       "DB_Bad_Konfig".Bad_Konfig[1].IO_Ein.WT_Einsetzen[1] := "FB_KP8_DB_1".KP8.Taste[6];
       "DB_Bad_Konfig".Bad_Konfig[1].IO_Ein.WT_Einsetzen[2] := "FB_KP8_DB_1".KP8.Taste[5];
       "DB_Bad_Konfig".Bad_Konfig[1].IO_Ein.WT_Einsetzen[3] := "FB_KP8_DB_1".KP8.Taste[4];
       "DB_Bad_Konfig".Bad_Konfig[1].IO_Ein.WT_Entnehmen[1] := "FB_KP8_DB_1".KP8.Taste[2];
       "DB_Bad_Konfig".Bad_Konfig[1].IO_Ein.WT_Entnehmen[2] := "FB_KP8_DB_1".KP8.Taste[1];
       "DB_Bad_Konfig".Bad_Konfig[1].IO_Ein.WT_Entnehmen[3] := "FB_KP8_DB_1".KP8.Taste[0];
       "DB_Bad_Konfig".Bad_Konfig[3].IO_Ein.WT_Einsetzen[1] := "FB_KP8_DB_2".KP8.Taste[6];
       "DB_Bad_Konfig".Bad_Konfig[3].IO_Ein.WT_Einsetzen[2] := "FB_KP8_DB_2".KP8.Taste[5];
       "DB_Bad_Konfig".Bad_Konfig[3].IO_Ein.WT_Einsetzen[3] := "FB_KP8_DB_2".KP8.Taste[4];
       "DB_Bad_Konfig".Bad_Konfig[3].IO_Ein.WT_Entnehmen[1] := "FB_KP8_DB_2".KP8.Taste[2];
       "DB_Bad_Konfig".Bad_Konfig[3].IO_Ein.WT_Entnehmen[2] := "FB_KP8_DB_2".KP8.Taste[1];
       "DB_Bad_Konfig".Bad_Konfig[3].IO_Ein.WT_Entnehmen[3] := "FB_KP8_DB_2".KP8.Taste[0];
       "DB_Bad_Konfig".Bad_Konfig[7].IO_Ein.WT_Einsetzen[1] := "FB_KP8_DB_4".KP8.Taste[6];
       "DB_Bad_Konfig".Bad_Konfig[7].IO_Ein.WT_Einsetzen[2] := "FB_KP8_DB_4".KP8.Taste[5];
       "DB_Bad_Konfig".Bad_Konfig[7].IO_Ein.WT_Einsetzen[3] := "FB_KP8_DB_4".KP8.Taste[4];
       "DB_Bad_Konfig".Bad_Konfig[7].IO_Ein.WT_Entnehmen[1] := "FB_KP8_DB_4".KP8.Taste[2];
       "DB_Bad_Konfig".Bad_Konfig[7].IO_Ein.WT_Entnehmen[2] := "FB_KP8_DB_4".KP8.Taste[1];
       "DB_Bad_Konfig".Bad_Konfig[7].IO_Ein.WT_Entnehmen[3] := "FB_KP8_DB_4".KP8.Taste[0];
       "DB_Bad_Konfig".Bad_Konfig[8].IO_Ein.WT_Einsetzen[1] := "FB_KP8_DB_5".KP8.Taste[6];
       "DB_Bad_Konfig".Bad_Konfig[8].IO_Ein.WT_Einsetzen[2] := "FB_KP8_DB_5".KP8.Taste[5];
       "DB_Bad_Konfig".Bad_Konfig[8].IO_Ein.WT_Einsetzen[3] := "FB_KP8_DB_5".KP8.Taste[4];
       "DB_Bad_Konfig".Bad_Konfig[8].IO_Ein.WT_Entnehmen[1] := "FB_KP8_DB_5".KP8.Taste[2];
       "DB_Bad_Konfig".Bad_Konfig[8].IO_Ein.WT_Entnehmen[2] := "FB_KP8_DB_5".KP8.Taste[1];
       "DB_Bad_Konfig".Bad_Konfig[8].IO_Ein.WT_Entnehmen[3] := "FB_KP8_DB_5".KP8.Taste[0];
       "DB_Bad_Konfig".Bad_Konfig[12].IO_Ein.WT_Einsetzen[1] := "FB_KP8_DB_7".KP8.Taste[6];
       "DB_Bad_Konfig".Bad_Konfig[12].IO_Ein.WT_Einsetzen[2] := "FB_KP8_DB_7".KP8.Taste[5];
       "DB_Bad_Konfig".Bad_Konfig[12].IO_Ein.WT_Einsetzen[3] := "FB_KP8_DB_7".KP8.Taste[4];
       "DB_Bad_Konfig".Bad_Konfig[12].IO_Ein.WT_Entnehmen[1] := "FB_KP8_DB_7".KP8.Taste[2];
       "DB_Bad_Konfig".Bad_Konfig[12].IO_Ein.WT_Entnehmen[2] := "FB_KP8_DB_7".KP8.Taste[1];
       "DB_Bad_Konfig".Bad_Konfig[12].IO_Ein.WT_Entnehmen[3] := "FB_KP8_DB_7".KP8.Taste[0];
       "DB_Bad_Konfig".Bad_Konfig[13].IO_Ein.WT_Einsetzen[1] := "FB_KP8_DB_8".KP8.Taste[6];
       "DB_Bad_Konfig".Bad_Konfig[13].IO_Ein.WT_Einsetzen[2] := "FB_KP8_DB_8".KP8.Taste[5];
       "DB_Bad_Konfig".Bad_Konfig[13].IO_Ein.WT_Einsetzen[3] := "FB_KP8_DB_8".KP8.Taste[4];
       "DB_Bad_Konfig".Bad_Konfig[13].IO_Ein.WT_Entnehmen[1] := "FB_KP8_DB_8".KP8.Taste[2];
       "DB_Bad_Konfig".Bad_Konfig[13].IO_Ein.WT_Entnehmen[2] := "FB_KP8_DB_8".KP8.Taste[1];
       "DB_Bad_Konfig".Bad_Konfig[13].IO_Ein.WT_Entnehmen[3] := "FB_KP8_DB_8".KP8.Taste[0];
       "DB_Bad_Konfig".Bad_Konfig[14].IO_Ein.WT_Einsetzen[1] := "FB_KP8_DB_9".KP8.Taste[6];
       "DB_Bad_Konfig".Bad_Konfig[14].IO_Ein.WT_Einsetzen[2] := "FB_KP8_DB_9".KP8.Taste[5];
       "DB_Bad_Konfig".Bad_Konfig[14].IO_Ein.WT_Einsetzen[3] := "FB_KP8_DB_9".KP8.Taste[4];
       "DB_Bad_Konfig".Bad_Konfig[14].IO_Ein.WT_Entnehmen[1] := "FB_KP8_DB_9".KP8.Taste[2];
       "DB_Bad_Konfig".Bad_Konfig[14].IO_Ein.WT_Entnehmen[2] := "FB_KP8_DB_9".KP8.Taste[1];
       "DB_Bad_Konfig".Bad_Konfig[14].IO_Ein.WT_Entnehmen[3] := "FB_KP8_DB_9".KP8.Taste[0];
       "DB_Bad_Konfig".Bad_Konfig[18].IO_Ein.WT_Einsetzen[1] := "FB_KP8_DB_11".KP8.Taste[6];
       "DB_Bad_Konfig".Bad_Konfig[18].IO_Ein.WT_Einsetzen[2] := "FB_KP8_DB_11".KP8.Taste[5];
       "DB_Bad_Konfig".Bad_Konfig[18].IO_Ein.WT_Einsetzen[3] := "FB_KP8_DB_11".KP8.Taste[4];
       "DB_Bad_Konfig".Bad_Konfig[18].IO_Ein.WT_Entnehmen[1] := "FB_KP8_DB_11".KP8.Taste[2];
       "DB_Bad_Konfig".Bad_Konfig[18].IO_Ein.WT_Entnehmen[2] := "FB_KP8_DB_11".KP8.Taste[1];
       "DB_Bad_Konfig".Bad_Konfig[18].IO_Ein.WT_Entnehmen[3] := "FB_KP8_DB_11".KP8.Taste[0];
       "DB_Bad_Konfig".Bad_Konfig[19].IO_Ein.WT_Einsetzen[1] := "FB_KP8_DB_12".KP8.Taste[6];
       "DB_Bad_Konfig".Bad_Konfig[19].IO_Ein.WT_Einsetzen[2] := "FB_KP8_DB_12".KP8.Taste[5];
       "DB_Bad_Konfig".Bad_Konfig[19].IO_Ein.WT_Einsetzen[3] := "FB_KP8_DB_12".KP8.Taste[4];
       "DB_Bad_Konfig".Bad_Konfig[19].IO_Ein.WT_Entnehmen[1] := "FB_KP8_DB_12".KP8.Taste[2];
       "DB_Bad_Konfig".Bad_Konfig[19].IO_Ein.WT_Entnehmen[2] := "FB_KP8_DB_12".KP8.Taste[1];
       "DB_Bad_Konfig".Bad_Konfig[19].IO_Ein.WT_Entnehmen[3] := "FB_KP8_DB_12".KP8.Taste[0];
       "DB_Bad_Konfig".Bad_Konfig[21].IO_Ein.WT_Einsetzen[1] := "FB_KP8_DB_13".KP8.Taste[6];
       "DB_Bad_Konfig".Bad_Konfig[21].IO_Ein.WT_Einsetzen[2] := "FB_KP8_DB_13".KP8.Taste[5];
       "DB_Bad_Konfig".Bad_Konfig[21].IO_Ein.WT_Einsetzen[3] := "FB_KP8_DB_13".KP8.Taste[4];
       "DB_Bad_Konfig".Bad_Konfig[21].IO_Ein.WT_Entnehmen[1] := "FB_KP8_DB_13".KP8.Taste[2];
       "DB_Bad_Konfig".Bad_Konfig[21].IO_Ein.WT_Entnehmen[2] := "FB_KP8_DB_13".KP8.Taste[1];
       "DB_Bad_Konfig".Bad_Konfig[21].IO_Ein.WT_Entnehmen[3] := "FB_KP8_DB_13".KP8.Taste[0];
       "DB_Bad_Konfig".Bad_Konfig[26].IO_Ein.WT_Einsetzen[1] := "FB_KP8_DB_15".KP8.Taste[6];
       "DB_Bad_Konfig".Bad_Konfig[26].IO_Ein.WT_Einsetzen[2] := "FB_KP8_DB_15".KP8.Taste[5];
       "DB_Bad_Konfig".Bad_Konfig[26].IO_Ein.WT_Einsetzen[3] := "FB_KP8_DB_15".KP8.Taste[4];
       "DB_Bad_Konfig".Bad_Konfig[26].IO_Ein.WT_Entnehmen[1] := "FB_KP8_DB_15".KP8.Taste[2];
       "DB_Bad_Konfig".Bad_Konfig[26].IO_Ein.WT_Entnehmen[2] := "FB_KP8_DB_15".KP8.Taste[1];
       "DB_Bad_Konfig".Bad_Konfig[26].IO_Ein.WT_Entnehmen[3] := "FB_KP8_DB_15".KP8.Taste[0];
       "DB_Bad_Konfig".Bad_Konfig[30].IO_Ein.WT_Einsetzen[1] := "FB_KP8_DB_17".KP8.Taste[6];
       "DB_Bad_Konfig".Bad_Konfig[30].IO_Ein.WT_Einsetzen[2] := "FB_KP8_DB_17".KP8.Taste[5];
       "DB_Bad_Konfig".Bad_Konfig[30].IO_Ein.WT_Einsetzen[3] := "FB_KP8_DB_17".KP8.Taste[4];
       "DB_Bad_Konfig".Bad_Konfig[30].IO_Ein.WT_Entnehmen[1] := "FB_KP8_DB_17".KP8.Taste[2];
       "DB_Bad_Konfig".Bad_Konfig[30].IO_Ein.WT_Entnehmen[2] := "FB_KP8_DB_17".KP8.Taste[1];
       "DB_Bad_Konfig".Bad_Konfig[30].IO_Ein.WT_Entnehmen[3] := "FB_KP8_DB_17".KP8.Taste[0];
       "DB_Bad_Konfig".Bad_Konfig[31].IO_Ein.WT_Einsetzen[1] := "FB_KP8_DB_18".KP8.Taste[6];
       "DB_Bad_Konfig".Bad_Konfig[31].IO_Ein.WT_Einsetzen[2] := "FB_KP8_DB_18".KP8.Taste[5];
       "DB_Bad_Konfig".Bad_Konfig[31].IO_Ein.WT_Einsetzen[3] := "FB_KP8_DB_18".KP8.Taste[4];
       "DB_Bad_Konfig".Bad_Konfig[31].IO_Ein.WT_Entnehmen[1] := "FB_KP8_DB_18".KP8.Taste[2];
       "DB_Bad_Konfig".Bad_Konfig[31].IO_Ein.WT_Entnehmen[2] := "FB_KP8_DB_18".KP8.Taste[1];
       "DB_Bad_Konfig".Bad_Konfig[31].IO_Ein.WT_Entnehmen[3] := "FB_KP8_DB_18".KP8.Taste[0];
       "DB_Bad_Konfig".Bad_Konfig[35].IO_Ein.WT_Einsetzen[1] := "FB_KP8_DB_20".KP8.Taste[6];
       "DB_Bad_Konfig".Bad_Konfig[35].IO_Ein.WT_Einsetzen[2] := "FB_KP8_DB_20".KP8.Taste[5];
       "DB_Bad_Konfig".Bad_Konfig[35].IO_Ein.WT_Einsetzen[3] := "FB_KP8_DB_20".KP8.Taste[4];
       "DB_Bad_Konfig".Bad_Konfig[35].IO_Ein.WT_Entnehmen[1] := "FB_KP8_DB_20".KP8.Taste[2];
       "DB_Bad_Konfig".Bad_Konfig[35].IO_Ein.WT_Entnehmen[2] := "FB_KP8_DB_20".KP8.Taste[1];
       "DB_Bad_Konfig".Bad_Konfig[35].IO_Ein.WT_Entnehmen[3] := "FB_KP8_DB_20".KP8.Taste[0];
       "DB_Bad_Konfig".Bad_Konfig[36].IO_Ein.WT_Einsetzen[1] := "FB_KP8_DB_21".KP8.Taste[6];
       "DB_Bad_Konfig".Bad_Konfig[36].IO_Ein.WT_Einsetzen[2] := "FB_KP8_DB_21".KP8.Taste[5];
       "DB_Bad_Konfig".Bad_Konfig[36].IO_Ein.WT_Einsetzen[3] := "FB_KP8_DB_21".KP8.Taste[4];
       "DB_Bad_Konfig".Bad_Konfig[36].IO_Ein.WT_Entnehmen[1] := "FB_KP8_DB_21".KP8.Taste[2];
       "DB_Bad_Konfig".Bad_Konfig[36].IO_Ein.WT_Entnehmen[2] := "FB_KP8_DB_21".KP8.Taste[1];
       "DB_Bad_Konfig".Bad_Konfig[36].IO_Ein.WT_Entnehmen[3] := "FB_KP8_DB_21".KP8.Taste[0];
       "DB_Bad_Konfig".Bad_Konfig[40].IO_Ein.WT_Einsetzen[1] := "FB_KP8_DB_23".KP8.Taste[6];
       "DB_Bad_Konfig".Bad_Konfig[40].IO_Ein.WT_Einsetzen[2] := "FB_KP8_DB_23".KP8.Taste[5];
       "DB_Bad_Konfig".Bad_Konfig[40].IO_Ein.WT_Einsetzen[3] := "FB_KP8_DB_23".KP8.Taste[4];
       "DB_Bad_Konfig".Bad_Konfig[40].IO_Ein.WT_Entnehmen[1] := "FB_KP8_DB_23".KP8.Taste[2];
       "DB_Bad_Konfig".Bad_Konfig[40].IO_Ein.WT_Entnehmen[2] := "FB_KP8_DB_23".KP8.Taste[1];
       "DB_Bad_Konfig".Bad_Konfig[40].IO_Ein.WT_Entnehmen[3] := "FB_KP8_DB_23".KP8.Taste[0];
       "DB_Bad_Konfig".Bad_Konfig[41].IO_Ein.WT_Einsetzen[1] := "FB_KP8_DB_24".KP8.Taste[6];
       "DB_Bad_Konfig".Bad_Konfig[41].IO_Ein.WT_Einsetzen[2] := "FB_KP8_DB_24".KP8.Taste[5];
       "DB_Bad_Konfig".Bad_Konfig[41].IO_Ein.WT_Einsetzen[3] := "FB_KP8_DB_24".KP8.Taste[4];
       "DB_Bad_Konfig".Bad_Konfig[41].IO_Ein.WT_Entnehmen[1] := "FB_KP8_DB_24".KP8.Taste[2];
       "DB_Bad_Konfig".Bad_Konfig[41].IO_Ein.WT_Entnehmen[2] := "FB_KP8_DB_24".KP8.Taste[1];
       "DB_Bad_Konfig".Bad_Konfig[41].IO_Ein.WT_Entnehmen[3] := "FB_KP8_DB_24".KP8.Taste[0];
       "DB_Bad_Konfig".Bad_Konfig[45].IO_Ein.WT_Einsetzen[1] := "FB_KP8_DB_26".KP8.Taste[6];
       "DB_Bad_Konfig".Bad_Konfig[45].IO_Ein.WT_Einsetzen[2] := "FB_KP8_DB_26".KP8.Taste[5];
       "DB_Bad_Konfig".Bad_Konfig[45].IO_Ein.WT_Einsetzen[3] := "FB_KP8_DB_26".KP8.Taste[4];
       "DB_Bad_Konfig".Bad_Konfig[45].IO_Ein.WT_Entnehmen[1] := "FB_KP8_DB_26".KP8.Taste[2];
       "DB_Bad_Konfig".Bad_Konfig[45].IO_Ein.WT_Entnehmen[2] := "FB_KP8_DB_26".KP8.Taste[1];
       "DB_Bad_Konfig".Bad_Konfig[45].IO_Ein.WT_Entnehmen[3] := "FB_KP8_DB_26".KP8.Taste[0];
       "DB_Bad_Konfig".Bad_Konfig[46].IO_Ein.WT_Einsetzen[1] := "FB_KP8_DB_27".KP8.Taste[6];
       "DB_Bad_Konfig".Bad_Konfig[46].IO_Ein.WT_Einsetzen[2] := "FB_KP8_DB_27".KP8.Taste[5];
       "DB_Bad_Konfig".Bad_Konfig[46].IO_Ein.WT_Einsetzen[3] := "FB_KP8_DB_27".KP8.Taste[4];
       "DB_Bad_Konfig".Bad_Konfig[46].IO_Ein.WT_Entnehmen[1] := "FB_KP8_DB_27".KP8.Taste[2];
       "DB_Bad_Konfig".Bad_Konfig[46].IO_Ein.WT_Entnehmen[2] := "FB_KP8_DB_27".KP8.Taste[1];
       "DB_Bad_Konfig".Bad_Konfig[46].IO_Ein.WT_Entnehmen[3] := "FB_KP8_DB_27".KP8.Taste[0];
       "DB_Bad_Konfig".Bad_Konfig[25].IO_Ein.WT_Einsetzen[1] := "FB_KP8_DB_28".KP8.Taste[6];
       "DB_Bad_Konfig".Bad_Konfig[25].IO_Ein.WT_Einsetzen[2] := "FB_KP8_DB_28".KP8.Taste[5];
       "DB_Bad_Konfig".Bad_Konfig[25].IO_Ein.WT_Einsetzen[3] := "FB_KP8_DB_28".KP8.Taste[4];
       "DB_Bad_Konfig".Bad_Konfig[25].IO_Ein.WT_Entnehmen[1] := "FB_KP8_DB_28".KP8.Taste[2];
       "DB_Bad_Konfig".Bad_Konfig[25].IO_Ein.WT_Entnehmen[2] := "FB_KP8_DB_28".KP8.Taste[1];
       "DB_Bad_Konfig".Bad_Konfig[25].IO_Ein.WT_Entnehmen[3] := "FB_KP8_DB_28".KP8.Taste[0];
       #pw := "DB_Bad_Konfig".Bad_Konfig[4].IO_Aus.Prio_Einsetzen_WT;
       IF (#pw >= 1) AND (#pw <= 3) THEN
           IF "FB_KP8_DB_3".KP8.Taste[4] THEN "DB_Bad_Konfig".Bad_Konfig[4].IO_Ein.WT_Einsetzen[#pw] := TRUE; END_IF;
       END_IF;
       #pw := "DB_Bad_Konfig".Bad_Konfig[4].IO_Aus.Prio_Entnehmen_WT;
       IF (#pw >= 1) AND (#pw <= 3) THEN
           IF "FB_KP8_DB_3".KP8.Taste[0] THEN "DB_Bad_Konfig".Bad_Konfig[4].IO_Ein.WT_Entnehmen[#pw] := TRUE; END_IF;
       END_IF;
       #pw := "DB_Bad_Konfig".Bad_Konfig[5].IO_Aus.Prio_Einsetzen_WT;
       IF (#pw >= 1) AND (#pw <= 3) THEN
           IF "FB_KP8_DB_3".KP8.Taste[5] THEN "DB_Bad_Konfig".Bad_Konfig[5].IO_Ein.WT_Einsetzen[#pw] := TRUE; END_IF;
       END_IF;
       #pw := "DB_Bad_Konfig".Bad_Konfig[5].IO_Aus.Prio_Entnehmen_WT;
       IF (#pw >= 1) AND (#pw <= 3) THEN
           IF "FB_KP8_DB_3".KP8.Taste[1] THEN "DB_Bad_Konfig".Bad_Konfig[5].IO_Ein.WT_Entnehmen[#pw] := TRUE; END_IF;
       END_IF;
       #pw := "DB_Bad_Konfig".Bad_Konfig[6].IO_Aus.Prio_Einsetzen_WT;
       IF (#pw >= 1) AND (#pw <= 3) THEN
           IF "FB_KP8_DB_3".KP8.Taste[6] THEN "DB_Bad_Konfig".Bad_Konfig[6].IO_Ein.WT_Einsetzen[#pw] := TRUE; END_IF;
       END_IF;
       #pw := "DB_Bad_Konfig".Bad_Konfig[6].IO_Aus.Prio_Entnehmen_WT;
       IF (#pw >= 1) AND (#pw <= 3) THEN
           IF "FB_KP8_DB_3".KP8.Taste[2] THEN "DB_Bad_Konfig".Bad_Konfig[6].IO_Ein.WT_Entnehmen[#pw] := TRUE; END_IF;
       END_IF;
       #pw := "DB_Bad_Konfig".Bad_Konfig[9].IO_Aus.Prio_Einsetzen_WT;
       IF (#pw >= 1) AND (#pw <= 3) THEN
           IF "FB_KP8_DB_6".KP8.Taste[4] THEN "DB_Bad_Konfig".Bad_Konfig[9].IO_Ein.WT_Einsetzen[#pw] := TRUE; END_IF;
       END_IF;
       #pw := "DB_Bad_Konfig".Bad_Konfig[9].IO_Aus.Prio_Entnehmen_WT;
       IF (#pw >= 1) AND (#pw <= 3) THEN
           IF "FB_KP8_DB_6".KP8.Taste[0] THEN "DB_Bad_Konfig".Bad_Konfig[9].IO_Ein.WT_Entnehmen[#pw] := TRUE; END_IF;
       END_IF;
       #pw := "DB_Bad_Konfig".Bad_Konfig[10].IO_Aus.Prio_Einsetzen_WT;
       IF (#pw >= 1) AND (#pw <= 3) THEN
           IF "FB_KP8_DB_6".KP8.Taste[5] THEN "DB_Bad_Konfig".Bad_Konfig[10].IO_Ein.WT_Einsetzen[#pw] := TRUE; END_IF;
       END_IF;
       #pw := "DB_Bad_Konfig".Bad_Konfig[10].IO_Aus.Prio_Entnehmen_WT;
       IF (#pw >= 1) AND (#pw <= 3) THEN
           IF "FB_KP8_DB_6".KP8.Taste[1] THEN "DB_Bad_Konfig".Bad_Konfig[10].IO_Ein.WT_Entnehmen[#pw] := TRUE; END_IF;
       END_IF;
       #pw := "DB_Bad_Konfig".Bad_Konfig[11].IO_Aus.Prio_Einsetzen_WT;
       IF (#pw >= 1) AND (#pw <= 3) THEN
           IF "FB_KP8_DB_6".KP8.Taste[6] THEN "DB_Bad_Konfig".Bad_Konfig[11].IO_Ein.WT_Einsetzen[#pw] := TRUE; END_IF;
       END_IF;
       #pw := "DB_Bad_Konfig".Bad_Konfig[11].IO_Aus.Prio_Entnehmen_WT;
       IF (#pw >= 1) AND (#pw <= 3) THEN
           IF "FB_KP8_DB_6".KP8.Taste[2] THEN "DB_Bad_Konfig".Bad_Konfig[11].IO_Ein.WT_Entnehmen[#pw] := TRUE; END_IF;
       END_IF;
       #pw := "DB_Bad_Konfig".Bad_Konfig[15].IO_Aus.Prio_Einsetzen_WT;
       IF (#pw >= 1) AND (#pw <= 3) THEN
           IF "FB_KP8_DB_10".KP8.Taste[4] THEN "DB_Bad_Konfig".Bad_Konfig[15].IO_Ein.WT_Einsetzen[#pw] := TRUE; END_IF;
       END_IF;
       #pw := "DB_Bad_Konfig".Bad_Konfig[15].IO_Aus.Prio_Entnehmen_WT;
       IF (#pw >= 1) AND (#pw <= 3) THEN
           IF "FB_KP8_DB_10".KP8.Taste[0] THEN "DB_Bad_Konfig".Bad_Konfig[15].IO_Ein.WT_Entnehmen[#pw] := TRUE; END_IF;
       END_IF;
       #pw := "DB_Bad_Konfig".Bad_Konfig[16].IO_Aus.Prio_Einsetzen_WT;
       IF (#pw >= 1) AND (#pw <= 3) THEN
           IF "FB_KP8_DB_10".KP8.Taste[5] THEN "DB_Bad_Konfig".Bad_Konfig[16].IO_Ein.WT_Einsetzen[#pw] := TRUE; END_IF;
       END_IF;
       #pw := "DB_Bad_Konfig".Bad_Konfig[16].IO_Aus.Prio_Entnehmen_WT;
       IF (#pw >= 1) AND (#pw <= 3) THEN
           IF "FB_KP8_DB_10".KP8.Taste[1] THEN "DB_Bad_Konfig".Bad_Konfig[16].IO_Ein.WT_Entnehmen[#pw] := TRUE; END_IF;
       END_IF;
       #pw := "DB_Bad_Konfig".Bad_Konfig[17].IO_Aus.Prio_Einsetzen_WT;
       IF (#pw >= 1) AND (#pw <= 3) THEN
           IF "FB_KP8_DB_10".KP8.Taste[6] THEN "DB_Bad_Konfig".Bad_Konfig[17].IO_Ein.WT_Einsetzen[#pw] := TRUE; END_IF;
       END_IF;
       #pw := "DB_Bad_Konfig".Bad_Konfig[17].IO_Aus.Prio_Entnehmen_WT;
       IF (#pw >= 1) AND (#pw <= 3) THEN
           IF "FB_KP8_DB_10".KP8.Taste[2] THEN "DB_Bad_Konfig".Bad_Konfig[17].IO_Ein.WT_Entnehmen[#pw] := TRUE; END_IF;
       END_IF;
       #pw := "DB_Bad_Konfig".Bad_Konfig[22].IO_Aus.Prio_Einsetzen_WT;
       IF (#pw >= 1) AND (#pw <= 3) THEN
           IF "FB_KP8_DB_14".KP8.Taste[4] THEN "DB_Bad_Konfig".Bad_Konfig[22].IO_Ein.WT_Einsetzen[#pw] := TRUE; END_IF;
       END_IF;
       #pw := "DB_Bad_Konfig".Bad_Konfig[22].IO_Aus.Prio_Entnehmen_WT;
       IF (#pw >= 1) AND (#pw <= 3) THEN
           IF "FB_KP8_DB_14".KP8.Taste[0] THEN "DB_Bad_Konfig".Bad_Konfig[22].IO_Ein.WT_Entnehmen[#pw] := TRUE; END_IF;
       END_IF;
       #pw := "DB_Bad_Konfig".Bad_Konfig[23].IO_Aus.Prio_Einsetzen_WT;
       IF (#pw >= 1) AND (#pw <= 3) THEN
           IF "FB_KP8_DB_14".KP8.Taste[5] THEN "DB_Bad_Konfig".Bad_Konfig[23].IO_Ein.WT_Einsetzen[#pw] := TRUE; END_IF;
       END_IF;
       #pw := "DB_Bad_Konfig".Bad_Konfig[23].IO_Aus.Prio_Entnehmen_WT;
       IF (#pw >= 1) AND (#pw <= 3) THEN
           IF "FB_KP8_DB_14".KP8.Taste[1] THEN "DB_Bad_Konfig".Bad_Konfig[23].IO_Ein.WT_Entnehmen[#pw] := TRUE; END_IF;
       END_IF;
       #pw := "DB_Bad_Konfig".Bad_Konfig[24].IO_Aus.Prio_Einsetzen_WT;
       IF (#pw >= 1) AND (#pw <= 3) THEN
           IF "FB_KP8_DB_14".KP8.Taste[6] THEN "DB_Bad_Konfig".Bad_Konfig[24].IO_Ein.WT_Einsetzen[#pw] := TRUE; END_IF;
       END_IF;
       #pw := "DB_Bad_Konfig".Bad_Konfig[24].IO_Aus.Prio_Entnehmen_WT;
       IF (#pw >= 1) AND (#pw <= 3) THEN
           IF "FB_KP8_DB_14".KP8.Taste[2] THEN "DB_Bad_Konfig".Bad_Konfig[24].IO_Ein.WT_Entnehmen[#pw] := TRUE; END_IF;
       END_IF;
       #pw := "DB_Bad_Konfig".Bad_Konfig[27].IO_Aus.Prio_Einsetzen_WT;
       IF (#pw >= 1) AND (#pw <= 3) THEN
           IF "FB_KP8_DB_16".KP8.Taste[4] THEN "DB_Bad_Konfig".Bad_Konfig[27].IO_Ein.WT_Einsetzen[#pw] := TRUE; END_IF;
       END_IF;
       #pw := "DB_Bad_Konfig".Bad_Konfig[27].IO_Aus.Prio_Entnehmen_WT;
       IF (#pw >= 1) AND (#pw <= 3) THEN
           IF "FB_KP8_DB_16".KP8.Taste[0] THEN "DB_Bad_Konfig".Bad_Konfig[27].IO_Ein.WT_Entnehmen[#pw] := TRUE; END_IF;
       END_IF;
       #pw := "DB_Bad_Konfig".Bad_Konfig[28].IO_Aus.Prio_Einsetzen_WT;
       IF (#pw >= 1) AND (#pw <= 3) THEN
           IF "FB_KP8_DB_16".KP8.Taste[5] THEN "DB_Bad_Konfig".Bad_Konfig[28].IO_Ein.WT_Einsetzen[#pw] := TRUE; END_IF;
       END_IF;
       #pw := "DB_Bad_Konfig".Bad_Konfig[28].IO_Aus.Prio_Entnehmen_WT;
       IF (#pw >= 1) AND (#pw <= 3) THEN
           IF "FB_KP8_DB_16".KP8.Taste[1] THEN "DB_Bad_Konfig".Bad_Konfig[28].IO_Ein.WT_Entnehmen[#pw] := TRUE; END_IF;
       END_IF;
       #pw := "DB_Bad_Konfig".Bad_Konfig[29].IO_Aus.Prio_Einsetzen_WT;
       IF (#pw >= 1) AND (#pw <= 3) THEN
           IF "FB_KP8_DB_16".KP8.Taste[6] THEN "DB_Bad_Konfig".Bad_Konfig[29].IO_Ein.WT_Einsetzen[#pw] := TRUE; END_IF;
       END_IF;
       #pw := "DB_Bad_Konfig".Bad_Konfig[29].IO_Aus.Prio_Entnehmen_WT;
       IF (#pw >= 1) AND (#pw <= 3) THEN
           IF "FB_KP8_DB_16".KP8.Taste[2] THEN "DB_Bad_Konfig".Bad_Konfig[29].IO_Ein.WT_Entnehmen[#pw] := TRUE; END_IF;
       END_IF;
       #pw := "DB_Bad_Konfig".Bad_Konfig[32].IO_Aus.Prio_Einsetzen_WT;
       IF (#pw >= 1) AND (#pw <= 3) THEN
           IF "FB_KP8_DB_19".KP8.Taste[4] THEN "DB_Bad_Konfig".Bad_Konfig[32].IO_Ein.WT_Einsetzen[#pw] := TRUE; END_IF;
       END_IF;
       #pw := "DB_Bad_Konfig".Bad_Konfig[32].IO_Aus.Prio_Entnehmen_WT;
       IF (#pw >= 1) AND (#pw <= 3) THEN
           IF "FB_KP8_DB_19".KP8.Taste[0] THEN "DB_Bad_Konfig".Bad_Konfig[32].IO_Ein.WT_Entnehmen[#pw] := TRUE; END_IF;
       END_IF;
       #pw := "DB_Bad_Konfig".Bad_Konfig[33].IO_Aus.Prio_Einsetzen_WT;
       IF (#pw >= 1) AND (#pw <= 3) THEN
           IF "FB_KP8_DB_19".KP8.Taste[5] THEN "DB_Bad_Konfig".Bad_Konfig[33].IO_Ein.WT_Einsetzen[#pw] := TRUE; END_IF;
       END_IF;
       #pw := "DB_Bad_Konfig".Bad_Konfig[33].IO_Aus.Prio_Entnehmen_WT;
       IF (#pw >= 1) AND (#pw <= 3) THEN
           IF "FB_KP8_DB_19".KP8.Taste[1] THEN "DB_Bad_Konfig".Bad_Konfig[33].IO_Ein.WT_Entnehmen[#pw] := TRUE; END_IF;
       END_IF;
       #pw := "DB_Bad_Konfig".Bad_Konfig[34].IO_Aus.Prio_Einsetzen_WT;
       IF (#pw >= 1) AND (#pw <= 3) THEN
           IF "FB_KP8_DB_19".KP8.Taste[6] THEN "DB_Bad_Konfig".Bad_Konfig[34].IO_Ein.WT_Einsetzen[#pw] := TRUE; END_IF;
       END_IF;
       #pw := "DB_Bad_Konfig".Bad_Konfig[34].IO_Aus.Prio_Entnehmen_WT;
       IF (#pw >= 1) AND (#pw <= 3) THEN
           IF "FB_KP8_DB_19".KP8.Taste[2] THEN "DB_Bad_Konfig".Bad_Konfig[34].IO_Ein.WT_Entnehmen[#pw] := TRUE; END_IF;
       END_IF;
       #pw := "DB_Bad_Konfig".Bad_Konfig[37].IO_Aus.Prio_Einsetzen_WT;
       IF (#pw >= 1) AND (#pw <= 3) THEN
           IF "FB_KP8_DB_22".KP8.Taste[4] THEN "DB_Bad_Konfig".Bad_Konfig[37].IO_Ein.WT_Einsetzen[#pw] := TRUE; END_IF;
       END_IF;
       #pw := "DB_Bad_Konfig".Bad_Konfig[37].IO_Aus.Prio_Entnehmen_WT;
       IF (#pw >= 1) AND (#pw <= 3) THEN
           IF "FB_KP8_DB_22".KP8.Taste[0] THEN "DB_Bad_Konfig".Bad_Konfig[37].IO_Ein.WT_Entnehmen[#pw] := TRUE; END_IF;
       END_IF;
       #pw := "DB_Bad_Konfig".Bad_Konfig[38].IO_Aus.Prio_Einsetzen_WT;
       IF (#pw >= 1) AND (#pw <= 3) THEN
           IF "FB_KP8_DB_22".KP8.Taste[5] THEN "DB_Bad_Konfig".Bad_Konfig[38].IO_Ein.WT_Einsetzen[#pw] := TRUE; END_IF;
       END_IF;
       #pw := "DB_Bad_Konfig".Bad_Konfig[38].IO_Aus.Prio_Entnehmen_WT;
       IF (#pw >= 1) AND (#pw <= 3) THEN
           IF "FB_KP8_DB_22".KP8.Taste[1] THEN "DB_Bad_Konfig".Bad_Konfig[38].IO_Ein.WT_Entnehmen[#pw] := TRUE; END_IF;
       END_IF;
       #pw := "DB_Bad_Konfig".Bad_Konfig[39].IO_Aus.Prio_Einsetzen_WT;
       IF (#pw >= 1) AND (#pw <= 3) THEN
           IF "FB_KP8_DB_22".KP8.Taste[6] THEN "DB_Bad_Konfig".Bad_Konfig[39].IO_Ein.WT_Einsetzen[#pw] := TRUE; END_IF;
       END_IF;
       #pw := "DB_Bad_Konfig".Bad_Konfig[39].IO_Aus.Prio_Entnehmen_WT;
       IF (#pw >= 1) AND (#pw <= 3) THEN
           IF "FB_KP8_DB_22".KP8.Taste[2] THEN "DB_Bad_Konfig".Bad_Konfig[39].IO_Ein.WT_Entnehmen[#pw] := TRUE; END_IF;
       END_IF;
       #pw := "DB_Bad_Konfig".Bad_Konfig[42].IO_Aus.Prio_Einsetzen_WT;
       IF (#pw >= 1) AND (#pw <= 3) THEN
           IF "FB_KP8_DB_25".KP8.Taste[4] THEN "DB_Bad_Konfig".Bad_Konfig[42].IO_Ein.WT_Einsetzen[#pw] := TRUE; END_IF;
       END_IF;
       #pw := "DB_Bad_Konfig".Bad_Konfig[42].IO_Aus.Prio_Entnehmen_WT;
       IF (#pw >= 1) AND (#pw <= 3) THEN
           IF "FB_KP8_DB_25".KP8.Taste[0] THEN "DB_Bad_Konfig".Bad_Konfig[42].IO_Ein.WT_Entnehmen[#pw] := TRUE; END_IF;
       END_IF;
       #pw := "DB_Bad_Konfig".Bad_Konfig[43].IO_Aus.Prio_Einsetzen_WT;
       IF (#pw >= 1) AND (#pw <= 3) THEN
           IF "FB_KP8_DB_25".KP8.Taste[5] THEN "DB_Bad_Konfig".Bad_Konfig[43].IO_Ein.WT_Einsetzen[#pw] := TRUE; END_IF;
       END_IF;
       #pw := "DB_Bad_Konfig".Bad_Konfig[43].IO_Aus.Prio_Entnehmen_WT;
       IF (#pw >= 1) AND (#pw <= 3) THEN
           IF "FB_KP8_DB_25".KP8.Taste[1] THEN "DB_Bad_Konfig".Bad_Konfig[43].IO_Ein.WT_Entnehmen[#pw] := TRUE; END_IF;
       END_IF;
       #pw := "DB_Bad_Konfig".Bad_Konfig[44].IO_Aus.Prio_Einsetzen_WT;
       IF (#pw >= 1) AND (#pw <= 3) THEN
           IF "FB_KP8_DB_25".KP8.Taste[6] THEN "DB_Bad_Konfig".Bad_Konfig[44].IO_Ein.WT_Einsetzen[#pw] := TRUE; END_IF;
       END_IF;
       #pw := "DB_Bad_Konfig".Bad_Konfig[44].IO_Aus.Prio_Entnehmen_WT;
       IF (#pw >= 1) AND (#pw <= 3) THEN
           IF "FB_KP8_DB_25".KP8.Taste[2] THEN "DB_Bad_Konfig".Bad_Konfig[44].IO_Ein.WT_Entnehmen[#pw] := TRUE; END_IF;
       END_IF;

       // Peripherie-Eingaenge
       "DB_Bad_Konfig".Bad_Konfig[7].IO_Ein.FI_Schutz_OK := "FI-Schutz 200F1 Heizung Bad 7 ist O.K.";
       "DB_Bad_Konfig".Bad_Konfig[7].IO_Ein.Kein_Uebertemp := "Heizung Bad 7 Keine uebertemperatur";
       "DB_Bad_Konfig".Bad_Konfig[7].IO_Ein.Niveau_OK := "Niveau Bad 7 OK";
       #rawWord := "Pt100 Heizung Bad 7"; #rawInt := WORD_TO_INT(#rawWord);
       "DB_Bad_Konfig".Bad_Konfig[7].IO_Ein.Ist_Temperatur_1 := INT_TO_REAL(#rawInt) / 10.0 + "DB_IPC_to_CPU".PT100_Offset[7];

       "DB_Bad_Konfig".Bad_Konfig[8].IO_Ein.FI_Schutz_OK := "FI-Schutz 210F1 Heizung Bad 8 ist O.K.";
       "DB_Bad_Konfig".Bad_Konfig[8].IO_Ein.Kein_Uebertemp := "Heizung Bad 8 Keine uebertemperatur";
       "DB_Bad_Konfig".Bad_Konfig[8].IO_Ein.Motorschutz_OK := "Motorschutz 215Q1 Pumpe Bad 8 ist O.K." AND "Wartungsschalter Pumpe Bad 8 ist eingeschaltet";
       "DB_Bad_Konfig".Bad_Konfig[8].IO_Ein.Niveau_OK := "Niveau Bad 8 OK";
       #rawWord := "Pt100 Heizung Bad 8"; #rawInt := WORD_TO_INT(#rawWord);
       "DB_Bad_Konfig".Bad_Konfig[8].IO_Ein.Ist_Temperatur_1 := INT_TO_REAL(#rawInt) / 10.0 + "DB_IPC_to_CPU".PT100_Offset[8];

       "DB_Bad_Konfig".Bad_Konfig[12].IO_Ein.FI_Schutz_OK := "FI-Schutz 220F1 Heizung Bad 12 ist O.K.";
       "DB_Bad_Konfig".Bad_Konfig[12].IO_Ein.Kein_Uebertemp := "Heizung Bad 12 Keine uebertemperatur";
       "DB_Bad_Konfig".Bad_Konfig[12].IO_Ein.Motorschutz_OK := "Motorschutz 225Q1 Pumpe Bad 12 ist O.K." AND "Wartungsschalter Pumpe Bad 12 ist eingeschaltet";
       "DB_Bad_Konfig".Bad_Konfig[12].IO_Ein.Niveau_OK := "Niveau Bad 12 OK";
       #rawWord := "Pt100 Heizung Bad 12"; #rawInt := WORD_TO_INT(#rawWord);
       "DB_Bad_Konfig".Bad_Konfig[12].IO_Ein.Ist_Temperatur_1 := INT_TO_REAL(#rawInt) / 10.0 + "DB_IPC_to_CPU".PT100_Offset[12];

       "DB_Bad_Konfig".Bad_Konfig[14].IO_Ein.Motorschutz_OK := "Motorschutz 235Q1 Pumpe Bad 14 ist O.K." AND "Wartungsschalter Pumpe Bad 14 ist eingeschaltet";
       "DB_Bad_Konfig".Bad_Konfig[18].IO_Ein.Motorschutz_OK := "Motorschutz 245Q1 Pumpe Bad 18 ist O.K." AND "Wartungsschalter Pumpe Bad 18 ist eingeschaltet";
       "DB_Bad_Konfig".Bad_Konfig[19].IO_Ein.Motorschutz_OK := "Motorschutz 255Q1 Pumpe Bad 19 ist O.K." AND "Wartungsschalter Pumpe Bad 19 ist eingeschaltet";
       "DB_Bad_Konfig".Bad_Konfig[21].IO_Ein.Motorschutz_OK := "Motorschutz 265Q1 Pumpe Bad 21 ist O.K." AND "Wartungsschalter Pumpe Bad 21 ist eingeschaltet";

       // Bad 25
       "DB_Bad_Konfig".Bad_Konfig[25].IO_Ein.FI_Schutz_OK := "Motorschutz und FI-Schutz 270Q1, 270F1 Heizung Bad 25 sind O.K." AND "Motorschutz und FI-Schutz 271Q1, 271F1 Heizung Bad 25 sind O.K.";
       "DB_Bad_Konfig".Bad_Konfig[25].IO_Ein.Kein_Uebertemp := "Heizung Bad 25 Keine uebertemperatur";
       "DB_Bad_Konfig".Bad_Konfig[25].IO_Ein.Motorschutz_OK := "Motorschutz 275Q1 Pumpe Bad 25 ist O.K." AND "Wartungsschalter Pumpe Bad 25 ist eingeschaltet";
       "DB_Bad_Konfig".Bad_Konfig[25].IO_Ein.Niveau_OK := "Niveau Bad 25 OK";
       "DB_Bad_Konfig".Bad_Konfig[25].IO_Ein.FU_Pumpe_Bereit := "FU Pumpe bereit";
       "DB_Bad_Konfig".Bad_Konfig[25].IO_Ein.FU_WB1_Bereit := "Warenbewegung 1 Bad 25 FU bereit";
       "DB_Bad_Konfig".Bad_Konfig[25].IO_Ein.FU_WB2_Bereit := "Warenbewegung 2 Bad 25 FU bereit";
       #rawWord := "Pt100 Heizung Bad 25"; #rawInt := WORD_TO_INT(#rawWord);
       "DB_Bad_Konfig".Bad_Konfig[25].IO_Ein.Ist_Temperatur_1 := INT_TO_REAL(#rawInt) / 10.0 + "DB_IPC_to_CPU".PT100_Offset[25];
       "DB_Bad_Konfig".Bad_Konfig[25].IO_Ein.Ist_Temperatur_2 := INT_TO_REAL(#rawInt) / 10.0 + "DB_IPC_to_CPU".PT100_Offset[25];

       "DB_Bad_Konfig".Bad_Konfig[26].IO_Ein.Motorschutz_OK := "Motorschutz 285Q1 Pumpe Bad 26 ist O.K." AND "Wartungsschalter Pumpe Bad 26 ist eingeschaltet";
       "DB_Bad_Konfig".Bad_Konfig[31].IO_Ein.Motorschutz_OK := "Motorschutz 295Q1 Pumpe Bad 31 ist O.K." AND "Wartungsschalter Pumpe Bad 31 ist eingeschaltet";

       "DB_Bad_Konfig".Bad_Konfig[36].IO_Ein.FI_Schutz_OK := "FI-Schutz 300F1 Heizung Bad 36 ist O.K.";
       "DB_Bad_Konfig".Bad_Konfig[36].IO_Ein.Kein_Uebertemp := "Heizung Bad 36 Keine uebertemperatur";
       "DB_Bad_Konfig".Bad_Konfig[36].IO_Ein.Niveau_OK := "Niveau Bad 36 OK";
       #rawWord := "Pt100 Heizung Bad 36"; #rawInt := WORD_TO_INT(#rawWord);
       "DB_Bad_Konfig".Bad_Konfig[36].IO_Ein.Ist_Temperatur_1 := INT_TO_REAL(#rawInt) / 10.0 + "DB_IPC_to_CPU".PT100_Offset[36];

       "DB_Bad_Konfig".Bad_Konfig[40].IO_Ein.FI_Schutz_OK := "FI-Schutz 310F1 Heizung Bad 40 ist O.K.";
       "DB_Bad_Konfig".Bad_Konfig[40].IO_Ein.Kein_Uebertemp := "Heizung Bad 40 Keine uebertemperatur";
       "DB_Bad_Konfig".Bad_Konfig[40].IO_Ein.Niveau_OK := "Niveau Bad 40 OK";
       #rawWord := "Pt100 Heizung Bad 40"; #rawInt := WORD_TO_INT(#rawWord);
       "DB_Bad_Konfig".Bad_Konfig[40].IO_Ein.Ist_Temperatur_1 := INT_TO_REAL(#rawInt) / 10.0 + "DB_IPC_to_CPU".PT100_Offset[40];

       "DB_Bad_Konfig".Bad_Konfig[41].IO_Ein.Motorschutz_OK := "Motorschutz 325Q1 Pumpe Bad 41 ist O.K." AND "Wartungsschalter Pumpe Bad 41 ist eingeschaltet";
       "DB_Bad_Konfig".Bad_Konfig[45].IO_Ein.Motorschutz_OK := "Motorschutz 335Q1 Pumpe Bad 45 ist O.K." AND "Wartungsschalter Pumpe Bad 45 ist eingeschaltet";

       "DB_Bad_Konfig".Bad_Konfig[46].IO_Ein.FI_Schutz_OK := "FI-Schutz 340F1 Heizung Bad 46 ist O.K.";
       "DB_Bad_Konfig".Bad_Konfig[46].IO_Ein.Kein_Uebertemp := "Heizung Bad 46 Keine uebertemperatur";
       "DB_Bad_Konfig".Bad_Konfig[46].IO_Ein.Niveau_OK := "Niveau Bad 46 OK";
       #rawWord := "Pt100 Heizung Bad 46"; #rawInt := WORD_TO_INT(#rawWord);
       "DB_Bad_Konfig".Bad_Konfig[46].IO_Ein.Ist_Temperatur_1 := INT_TO_REAL(#rawInt) / 10.0 + "DB_IPC_to_CPU".PT100_Offset[46];

   ELSIF #Richtung = 2 THEN
       "FB_KP8_DB_1".KP8.DO[4] := "DB_Bad_Konfig".Bad_Konfig[1].IO_Aus.Ampel_Orange;
       "FB_KP8_DB_1".KP8.DO[5] := "DB_Bad_Konfig".Bad_Konfig[1].IO_Aus.Ampel_Gruen;
       "FB_KP8_DB_1".KP8.DO[6] := "DB_Bad_Konfig".Bad_Konfig[1].IO_Aus.Ampel_Rot;
       "FB_KP8_DB_2".KP8.DO[4] := "DB_Bad_Konfig".Bad_Konfig[3].IO_Aus.Ampel_Orange;
       "FB_KP8_DB_2".KP8.DO[5] := "DB_Bad_Konfig".Bad_Konfig[3].IO_Aus.Ampel_Gruen;
       "FB_KP8_DB_2".KP8.DO[6] := "DB_Bad_Konfig".Bad_Konfig[3].IO_Aus.Ampel_Rot;
       "FB_KP8_DB_4".KP8.DO[4] := "DB_Bad_Konfig".Bad_Konfig[7].IO_Aus.Ampel_Orange;
       "FB_KP8_DB_4".KP8.DO[5] := "DB_Bad_Konfig".Bad_Konfig[7].IO_Aus.Ampel_Gruen;
       "FB_KP8_DB_4".KP8.DO[6] := "DB_Bad_Konfig".Bad_Konfig[7].IO_Aus.Ampel_Rot;
       "FB_KP8_DB_5".KP8.DO[4] := "DB_Bad_Konfig".Bad_Konfig[8].IO_Aus.Ampel_Orange;
       "FB_KP8_DB_5".KP8.DO[5] := "DB_Bad_Konfig".Bad_Konfig[8].IO_Aus.Ampel_Gruen;
       "FB_KP8_DB_5".KP8.DO[6] := "DB_Bad_Konfig".Bad_Konfig[8].IO_Aus.Ampel_Rot;
       "FB_KP8_DB_7".KP8.DO[4] := "DB_Bad_Konfig".Bad_Konfig[12].IO_Aus.Ampel_Orange;
       "FB_KP8_DB_7".KP8.DO[5] := "DB_Bad_Konfig".Bad_Konfig[12].IO_Aus.Ampel_Gruen;
       "FB_KP8_DB_7".KP8.DO[6] := "DB_Bad_Konfig".Bad_Konfig[12].IO_Aus.Ampel_Rot;
       "FB_KP8_DB_8".KP8.DO[4] := "DB_Bad_Konfig".Bad_Konfig[13].IO_Aus.Ampel_Orange;
       "FB_KP8_DB_8".KP8.DO[5] := "DB_Bad_Konfig".Bad_Konfig[13].IO_Aus.Ampel_Gruen;
       "FB_KP8_DB_8".KP8.DO[6] := "DB_Bad_Konfig".Bad_Konfig[13].IO_Aus.Ampel_Rot;
       "FB_KP8_DB_9".KP8.DO[4] := "DB_Bad_Konfig".Bad_Konfig[14].IO_Aus.Ampel_Orange;
       "FB_KP8_DB_9".KP8.DO[5] := "DB_Bad_Konfig".Bad_Konfig[14].IO_Aus.Ampel_Gruen;
       "FB_KP8_DB_9".KP8.DO[6] := "DB_Bad_Konfig".Bad_Konfig[14].IO_Aus.Ampel_Rot;
       "FB_KP8_DB_11".KP8.DO[4] := "DB_Bad_Konfig".Bad_Konfig[18].IO_Aus.Ampel_Orange;
       "FB_KP8_DB_11".KP8.DO[5] := "DB_Bad_Konfig".Bad_Konfig[18].IO_Aus.Ampel_Gruen;
       "FB_KP8_DB_11".KP8.DO[6] := "DB_Bad_Konfig".Bad_Konfig[18].IO_Aus.Ampel_Rot;
       "FB_KP8_DB_12".KP8.DO[4] := "DB_Bad_Konfig".Bad_Konfig[19].IO_Aus.Ampel_Orange;
       "FB_KP8_DB_12".KP8.DO[5] := "DB_Bad_Konfig".Bad_Konfig[19].IO_Aus.Ampel_Gruen;
       "FB_KP8_DB_12".KP8.DO[6] := "DB_Bad_Konfig".Bad_Konfig[19].IO_Aus.Ampel_Rot;
       "FB_KP8_DB_13".KP8.DO[4] := "DB_Bad_Konfig".Bad_Konfig[21].IO_Aus.Ampel_Orange;
       "FB_KP8_DB_13".KP8.DO[5] := "DB_Bad_Konfig".Bad_Konfig[21].IO_Aus.Ampel_Gruen;
       "FB_KP8_DB_13".KP8.DO[6] := "DB_Bad_Konfig".Bad_Konfig[21].IO_Aus.Ampel_Rot;
       "FB_KP8_DB_15".KP8.DO[4] := "DB_Bad_Konfig".Bad_Konfig[26].IO_Aus.Ampel_Orange;
       "FB_KP8_DB_15".KP8.DO[5] := "DB_Bad_Konfig".Bad_Konfig[26].IO_Aus.Ampel_Gruen;
       "FB_KP8_DB_15".KP8.DO[6] := "DB_Bad_Konfig".Bad_Konfig[26].IO_Aus.Ampel_Rot;
       "FB_KP8_DB_17".KP8.DO[4] := "DB_Bad_Konfig".Bad_Konfig[30].IO_Aus.Ampel_Orange;
       "FB_KP8_DB_17".KP8.DO[5] := "DB_Bad_Konfig".Bad_Konfig[30].IO_Aus.Ampel_Gruen;
       "FB_KP8_DB_17".KP8.DO[6] := "DB_Bad_Konfig".Bad_Konfig[30].IO_Aus.Ampel_Rot;
       "FB_KP8_DB_18".KP8.DO[4] := "DB_Bad_Konfig".Bad_Konfig[31].IO_Aus.Ampel_Orange;
       "FB_KP8_DB_18".KP8.DO[5] := "DB_Bad_Konfig".Bad_Konfig[31].IO_Aus.Ampel_Gruen;
       "FB_KP8_DB_18".KP8.DO[6] := "DB_Bad_Konfig".Bad_Konfig[31].IO_Aus.Ampel_Rot;
       "FB_KP8_DB_20".KP8.DO[4] := "DB_Bad_Konfig".Bad_Konfig[35].IO_Aus.Ampel_Orange;
       "FB_KP8_DB_20".KP8.DO[5] := "DB_Bad_Konfig".Bad_Konfig[35].IO_Aus.Ampel_Gruen;
       "FB_KP8_DB_20".KP8.DO[6] := "DB_Bad_Konfig".Bad_Konfig[35].IO_Aus.Ampel_Rot;
       "FB_KP8_DB_21".KP8.DO[4] := "DB_Bad_Konfig".Bad_Konfig[36].IO_Aus.Ampel_Orange;
       "FB_KP8_DB_21".KP8.DO[5] := "DB_Bad_Konfig".Bad_Konfig[36].IO_Aus.Ampel_Gruen;
       "FB_KP8_DB_21".KP8.DO[6] := "DB_Bad_Konfig".Bad_Konfig[36].IO_Aus.Ampel_Rot;
       "FB_KP8_DB_23".KP8.DO[4] := "DB_Bad_Konfig".Bad_Konfig[40].IO_Aus.Ampel_Orange;
       "FB_KP8_DB_23".KP8.DO[5] := "DB_Bad_Konfig".Bad_Konfig[40].IO_Aus.Ampel_Gruen;
       "FB_KP8_DB_23".KP8.DO[6] := "DB_Bad_Konfig".Bad_Konfig[40].IO_Aus.Ampel_Rot;
       "FB_KP8_DB_24".KP8.DO[4] := "DB_Bad_Konfig".Bad_Konfig[41].IO_Aus.Ampel_Orange;
       "FB_KP8_DB_24".KP8.DO[5] := "DB_Bad_Konfig".Bad_Konfig[41].IO_Aus.Ampel_Gruen;
       "FB_KP8_DB_24".KP8.DO[6] := "DB_Bad_Konfig".Bad_Konfig[41].IO_Aus.Ampel_Rot;
       "FB_KP8_DB_26".KP8.DO[4] := "DB_Bad_Konfig".Bad_Konfig[45].IO_Aus.Ampel_Orange;
       "FB_KP8_DB_26".KP8.DO[5] := "DB_Bad_Konfig".Bad_Konfig[45].IO_Aus.Ampel_Gruen;
       "FB_KP8_DB_26".KP8.DO[6] := "DB_Bad_Konfig".Bad_Konfig[45].IO_Aus.Ampel_Rot;
       "FB_KP8_DB_27".KP8.DO[4] := "DB_Bad_Konfig".Bad_Konfig[46].IO_Aus.Ampel_Orange;
       "FB_KP8_DB_27".KP8.DO[5] := "DB_Bad_Konfig".Bad_Konfig[46].IO_Aus.Ampel_Gruen;
       "FB_KP8_DB_27".KP8.DO[6] := "DB_Bad_Konfig".Bad_Konfig[46].IO_Aus.Ampel_Rot;
       "FB_KP8_DB_28".KP8.DO[4] := "DB_Bad_Konfig".Bad_Konfig[25].IO_Aus.Ampel_Orange;
       "FB_KP8_DB_28".KP8.DO[5] := "DB_Bad_Konfig".Bad_Konfig[25].IO_Aus.Ampel_Gruen;
       "FB_KP8_DB_28".KP8.DO[6] := "DB_Bad_Konfig".Bad_Konfig[25].IO_Aus.Ampel_Rot;
       "FB_KP8_DB_3".KP8.DO[4] := "DB_Bad_Konfig".Bad_Konfig[4].IO_Aus.Ampel_Orange OR "DB_Bad_Konfig".Bad_Konfig[5].IO_Aus.Ampel_Orange OR "DB_Bad_Konfig".Bad_Konfig[6].IO_Aus.Ampel_Orange;
       "FB_KP8_DB_3".KP8.DO[5] := "DB_Bad_Konfig".Bad_Konfig[4].IO_Aus.Ampel_Gruen OR "DB_Bad_Konfig".Bad_Konfig[5].IO_Aus.Ampel_Gruen OR "DB_Bad_Konfig".Bad_Konfig[6].IO_Aus.Ampel_Gruen;
       "FB_KP8_DB_3".KP8.DO[6] := "DB_Bad_Konfig".Bad_Konfig[4].IO_Aus.Ampel_Rot OR "DB_Bad_Konfig".Bad_Konfig[5].IO_Aus.Ampel_Rot OR "DB_Bad_Konfig".Bad_Konfig[6].IO_Aus.Ampel_Rot;
       "FB_KP8_DB_6".KP8.DO[4] := "DB_Bad_Konfig".Bad_Konfig[9].IO_Aus.Ampel_Orange OR "DB_Bad_Konfig".Bad_Konfig[10].IO_Aus.Ampel_Orange OR "DB_Bad_Konfig".Bad_Konfig[11].IO_Aus.Ampel_Orange;
       "FB_KP8_DB_6".KP8.DO[5] := "DB_Bad_Konfig".Bad_Konfig[9].IO_Aus.Ampel_Gruen OR "DB_Bad_Konfig".Bad_Konfig[10].IO_Aus.Ampel_Gruen OR "DB_Bad_Konfig".Bad_Konfig[11].IO_Aus.Ampel_Gruen;
       "FB_KP8_DB_6".KP8.DO[6] := "DB_Bad_Konfig".Bad_Konfig[9].IO_Aus.Ampel_Rot OR "DB_Bad_Konfig".Bad_Konfig[10].IO_Aus.Ampel_Rot OR "DB_Bad_Konfig".Bad_Konfig[11].IO_Aus.Ampel_Rot;
       "FB_KP8_DB_10".KP8.DO[4] := "DB_Bad_Konfig".Bad_Konfig[15].IO_Aus.Ampel_Orange OR "DB_Bad_Konfig".Bad_Konfig[16].IO_Aus.Ampel_Orange OR "DB_Bad_Konfig".Bad_Konfig[17].IO_Aus.Ampel_Orange;
       "FB_KP8_DB_10".KP8.DO[5] := "DB_Bad_Konfig".Bad_Konfig[15].IO_Aus.Ampel_Gruen OR "DB_Bad_Konfig".Bad_Konfig[16].IO_Aus.Ampel_Gruen OR "DB_Bad_Konfig".Bad_Konfig[17].IO_Aus.Ampel_Gruen;
       "FB_KP8_DB_10".KP8.DO[6] := "DB_Bad_Konfig".Bad_Konfig[15].IO_Aus.Ampel_Rot OR "DB_Bad_Konfig".Bad_Konfig[16].IO_Aus.Ampel_Rot OR "DB_Bad_Konfig".Bad_Konfig[17].IO_Aus.Ampel_Rot;
       "FB_KP8_DB_14".KP8.DO[4] := "DB_Bad_Konfig".Bad_Konfig[22].IO_Aus.Ampel_Orange OR "DB_Bad_Konfig".Bad_Konfig[23].IO_Aus.Ampel_Orange OR "DB_Bad_Konfig".Bad_Konfig[24].IO_Aus.Ampel_Orange;
       "FB_KP8_DB_14".KP8.DO[5] := "DB_Bad_Konfig".Bad_Konfig[22].IO_Aus.Ampel_Gruen OR "DB_Bad_Konfig".Bad_Konfig[23].IO_Aus.Ampel_Gruen OR "DB_Bad_Konfig".Bad_Konfig[24].IO_Aus.Ampel_Gruen;
       "FB_KP8_DB_14".KP8.DO[6] := "DB_Bad_Konfig".Bad_Konfig[22].IO_Aus.Ampel_Rot OR "DB_Bad_Konfig".Bad_Konfig[23].IO_Aus.Ampel_Rot OR "DB_Bad_Konfig".Bad_Konfig[24].IO_Aus.Ampel_Rot;
       "FB_KP8_DB_16".KP8.DO[4] := "DB_Bad_Konfig".Bad_Konfig[27].IO_Aus.Ampel_Orange OR "DB_Bad_Konfig".Bad_Konfig[28].IO_Aus.Ampel_Orange OR "DB_Bad_Konfig".Bad_Konfig[29].IO_Aus.Ampel_Orange;
       "FB_KP8_DB_16".KP8.DO[5] := "DB_Bad_Konfig".Bad_Konfig[27].IO_Aus.Ampel_Gruen OR "DB_Bad_Konfig".Bad_Konfig[28].IO_Aus.Ampel_Gruen OR "DB_Bad_Konfig".Bad_Konfig[29].IO_Aus.Ampel_Gruen;
       "FB_KP8_DB_16".KP8.DO[6] := "DB_Bad_Konfig".Bad_Konfig[27].IO_Aus.Ampel_Rot OR "DB_Bad_Konfig".Bad_Konfig[28].IO_Aus.Ampel_Rot OR "DB_Bad_Konfig".Bad_Konfig[29].IO_Aus.Ampel_Rot;
       "FB_KP8_DB_19".KP8.DO[4] := "DB_Bad_Konfig".Bad_Konfig[32].IO_Aus.Ampel_Orange OR "DB_Bad_Konfig".Bad_Konfig[33].IO_Aus.Ampel_Orange OR "DB_Bad_Konfig".Bad_Konfig[34].IO_Aus.Ampel_Orange;
       "FB_KP8_DB_19".KP8.DO[5] := "DB_Bad_Konfig".Bad_Konfig[32].IO_Aus.Ampel_Gruen OR "DB_Bad_Konfig".Bad_Konfig[33].IO_Aus.Ampel_Gruen OR "DB_Bad_Konfig".Bad_Konfig[34].IO_Aus.Ampel_Gruen;
       "FB_KP8_DB_19".KP8.DO[6] := "DB_Bad_Konfig".Bad_Konfig[32].IO_Aus.Ampel_Rot OR "DB_Bad_Konfig".Bad_Konfig[33].IO_Aus.Ampel_Rot OR "DB_Bad_Konfig".Bad_Konfig[34].IO_Aus.Ampel_Rot;
       "FB_KP8_DB_22".KP8.DO[4] := "DB_Bad_Konfig".Bad_Konfig[37].IO_Aus.Ampel_Orange OR "DB_Bad_Konfig".Bad_Konfig[38].IO_Aus.Ampel_Orange OR "DB_Bad_Konfig".Bad_Konfig[39].IO_Aus.Ampel_Orange;
       "FB_KP8_DB_22".KP8.DO[5] := "DB_Bad_Konfig".Bad_Konfig[37].IO_Aus.Ampel_Gruen OR "DB_Bad_Konfig".Bad_Konfig[38].IO_Aus.Ampel_Gruen OR "DB_Bad_Konfig".Bad_Konfig[39].IO_Aus.Ampel_Gruen;
       "FB_KP8_DB_22".KP8.DO[6] := "DB_Bad_Konfig".Bad_Konfig[37].IO_Aus.Ampel_Rot OR "DB_Bad_Konfig".Bad_Konfig[38].IO_Aus.Ampel_Rot OR "DB_Bad_Konfig".Bad_Konfig[39].IO_Aus.Ampel_Rot;
       "FB_KP8_DB_25".KP8.DO[4] := "DB_Bad_Konfig".Bad_Konfig[42].IO_Aus.Ampel_Orange OR "DB_Bad_Konfig".Bad_Konfig[43].IO_Aus.Ampel_Orange OR "DB_Bad_Konfig".Bad_Konfig[44].IO_Aus.Ampel_Orange;
       "FB_KP8_DB_25".KP8.DO[5] := "DB_Bad_Konfig".Bad_Konfig[42].IO_Aus.Ampel_Gruen OR "DB_Bad_Konfig".Bad_Konfig[43].IO_Aus.Ampel_Gruen OR "DB_Bad_Konfig".Bad_Konfig[44].IO_Aus.Ampel_Gruen;
       "FB_KP8_DB_25".KP8.DO[6] := "DB_Bad_Konfig".Bad_Konfig[42].IO_Aus.Ampel_Rot OR "DB_Bad_Konfig".Bad_Konfig[43].IO_Aus.Ampel_Rot OR "DB_Bad_Konfig".Bad_Konfig[44].IO_Aus.Ampel_Rot;

       // KP8 Tasten-LEDs
       IF "DB_Bad_Konfig".Bad_Konfig[1].IO_Aus.LED_Einsetzen[1] THEN "FB_KP8_DB_1".KP8.LED[6] := 5; ELSE "FB_KP8_DB_1".KP8.LED[6] := 0; END_IF;
       IF "DB_Bad_Konfig".Bad_Konfig[1].IO_Aus.LED_Entnehmen[1] THEN
           IF "DB_Bad_Konfig".Bad_Konfig[1].IO_Aus.LED_Vorwarn[1] THEN "FB_KP8_DB_1".KP8.LED[2] := 4; ELSE "FB_KP8_DB_1".KP8.LED[2] := 5; END_IF;
       ELSE "FB_KP8_DB_1".KP8.LED[2] := 0; END_IF;
       IF "DB_Bad_Konfig".Bad_Konfig[1].IO_Aus.LED_Einsetzen[2] THEN "FB_KP8_DB_1".KP8.LED[5] := 5; ELSE "FB_KP8_DB_1".KP8.LED[5] := 0; END_IF;
       IF "DB_Bad_Konfig".Bad_Konfig[1].IO_Aus.LED_Entnehmen[2] THEN
           IF "DB_Bad_Konfig".Bad_Konfig[1].IO_Aus.LED_Vorwarn[2] THEN "FB_KP8_DB_1".KP8.LED[1] := 4; ELSE "FB_KP8_DB_1".KP8.LED[1] := 5; END_IF;
       ELSE "FB_KP8_DB_1".KP8.LED[1] := 0; END_IF;
       IF "DB_Bad_Konfig".Bad_Konfig[1].IO_Aus.LED_Einsetzen[3] THEN "FB_KP8_DB_1".KP8.LED[4] := 5; ELSE "FB_KP8_DB_1".KP8.LED[4] := 0; END_IF;
       IF "DB_Bad_Konfig".Bad_Konfig[1].IO_Aus.LED_Entnehmen[3] THEN
           IF "DB_Bad_Konfig".Bad_Konfig[1].IO_Aus.LED_Vorwarn[3] THEN "FB_KP8_DB_1".KP8.LED[0] := 4; ELSE "FB_KP8_DB_1".KP8.LED[0] := 5; END_IF;
       ELSE "FB_KP8_DB_1".KP8.LED[0] := 0; END_IF;
       IF "DB_Bad_Konfig".Bad_Konfig[1].IO_Aus.LED_Heizung_Aktiv THEN "FB_KP8_DB_1".KP8.LED[3] := 4; ELSE "FB_KP8_DB_1".KP8.LED[3] := 0; END_IF;
       IF "DB_Bad_Konfig".Bad_Konfig[1].IO_Aus.LED_Stoerung THEN "FB_KP8_DB_1".KP8.LED[7] := 1; ELSE "FB_KP8_DB_1".KP8.LED[7] := 0; END_IF;
       IF "DB_Bad_Konfig".Bad_Konfig[3].IO_Aus.LED_Einsetzen[1] THEN "FB_KP8_DB_2".KP8.LED[6] := 5; ELSE "FB_KP8_DB_2".KP8.LED[6] := 0; END_IF;
       IF "DB_Bad_Konfig".Bad_Konfig[3].IO_Aus.LED_Entnehmen[1] THEN
           IF "DB_Bad_Konfig".Bad_Konfig[3].IO_Aus.LED_Vorwarn[1] THEN "FB_KP8_DB_2".KP8.LED[2] := 4; ELSE "FB_KP8_DB_2".KP8.LED[2] := 5; END_IF;
       ELSE "FB_KP8_DB_2".KP8.LED[2] := 0; END_IF;
       IF "DB_Bad_Konfig".Bad_Konfig[3].IO_Aus.LED_Einsetzen[2] THEN "FB_KP8_DB_2".KP8.LED[5] := 5; ELSE "FB_KP8_DB_2".KP8.LED[5] := 0; END_IF;
       IF "DB_Bad_Konfig".Bad_Konfig[3].IO_Aus.LED_Entnehmen[2] THEN
           IF "DB_Bad_Konfig".Bad_Konfig[3].IO_Aus.LED_Vorwarn[2] THEN "FB_KP8_DB_2".KP8.LED[1] := 4; ELSE "FB_KP8_DB_2".KP8.LED[1] := 5; END_IF;
       ELSE "FB_KP8_DB_2".KP8.LED[1] := 0; END_IF;
       IF "DB_Bad_Konfig".Bad_Konfig[3].IO_Aus.LED_Einsetzen[3] THEN "FB_KP8_DB_2".KP8.LED[4] := 5; ELSE "FB_KP8_DB_2".KP8.LED[4] := 0; END_IF;
       IF "DB_Bad_Konfig".Bad_Konfig[3].IO_Aus.LED_Entnehmen[3] THEN
           IF "DB_Bad_Konfig".Bad_Konfig[3].IO_Aus.LED_Vorwarn[3] THEN "FB_KP8_DB_2".KP8.LED[0] := 4; ELSE "FB_KP8_DB_2".KP8.LED[0] := 5; END_IF;
       ELSE "FB_KP8_DB_2".KP8.LED[0] := 0; END_IF;
       IF "DB_Bad_Konfig".Bad_Konfig[3].IO_Aus.LED_Heizung_Aktiv THEN "FB_KP8_DB_2".KP8.LED[3] := 4; ELSE "FB_KP8_DB_2".KP8.LED[3] := 0; END_IF;
       IF "DB_Bad_Konfig".Bad_Konfig[3].IO_Aus.LED_Stoerung THEN "FB_KP8_DB_2".KP8.LED[7] := 1; ELSE "FB_KP8_DB_2".KP8.LED[7] := 0; END_IF;
       IF "DB_Bad_Konfig".Bad_Konfig[7].IO_Aus.LED_Einsetzen[1] THEN "FB_KP8_DB_4".KP8.LED[6] := 5; ELSE "FB_KP8_DB_4".KP8.LED[6] := 0; END_IF;
       IF "DB_Bad_Konfig".Bad_Konfig[7].IO_Aus.LED_Entnehmen[1] THEN
           IF "DB_Bad_Konfig".Bad_Konfig[7].IO_Aus.LED_Vorwarn[1] THEN "FB_KP8_DB_4".KP8.LED[2] := 4; ELSE "FB_KP8_DB_4".KP8.LED[2] := 5; END_IF;
       ELSE "FB_KP8_DB_4".KP8.LED[2] := 0; END_IF;
       IF "DB_Bad_Konfig".Bad_Konfig[7].IO_Aus.LED_Einsetzen[2] THEN "FB_KP8_DB_4".KP8.LED[5] := 5; ELSE "FB_KP8_DB_4".KP8.LED[5] := 0; END_IF;
       IF "DB_Bad_Konfig".Bad_Konfig[7].IO_Aus.LED_Entnehmen[2] THEN
           IF "DB_Bad_Konfig".Bad_Konfig[7].IO_Aus.LED_Vorwarn[2] THEN "FB_KP8_DB_4".KP8.LED[1] := 4; ELSE "FB_KP8_DB_4".KP8.LED[1] := 5; END_IF;
       ELSE "FB_KP8_DB_4".KP8.LED[1] := 0; END_IF;
       IF "DB_Bad_Konfig".Bad_Konfig[7].IO_Aus.LED_Einsetzen[3] THEN "FB_KP8_DB_4".KP8.LED[4] := 5; ELSE "FB_KP8_DB_4".KP8.LED[4] := 0; END_IF;
       IF "DB_Bad_Konfig".Bad_Konfig[7].IO_Aus.LED_Entnehmen[3] THEN
           IF "DB_Bad_Konfig".Bad_Konfig[7].IO_Aus.LED_Vorwarn[3] THEN "FB_KP8_DB_4".KP8.LED[0] := 4; ELSE "FB_KP8_DB_4".KP8.LED[0] := 5; END_IF;
       ELSE "FB_KP8_DB_4".KP8.LED[0] := 0; END_IF;
       IF "DB_Bad_Konfig".Bad_Konfig[7].IO_Aus.LED_Heizung_Aktiv THEN "FB_KP8_DB_4".KP8.LED[3] := 4; ELSE "FB_KP8_DB_4".KP8.LED[3] := 0; END_IF;
       IF "DB_Bad_Konfig".Bad_Konfig[7].IO_Aus.LED_Stoerung THEN "FB_KP8_DB_4".KP8.LED[7] := 1; ELSE "FB_KP8_DB_4".KP8.LED[7] := 0; END_IF;
       IF "DB_Bad_Konfig".Bad_Konfig[8].IO_Aus.LED_Einsetzen[1] THEN "FB_KP8_DB_5".KP8.LED[6] := 5; ELSE "FB_KP8_DB_5".KP8.LED[6] := 0; END_IF;
       IF "DB_Bad_Konfig".Bad_Konfig[8].IO_Aus.LED_Entnehmen[1] THEN
           IF "DB_Bad_Konfig".Bad_Konfig[8].IO_Aus.LED_Vorwarn[1] THEN "FB_KP8_DB_5".KP8.LED[2] := 4; ELSE "FB_KP8_DB_5".KP8.LED[2] := 5; END_IF;
       ELSE "FB_KP8_DB_5".KP8.LED[2] := 0; END_IF;
       IF "DB_Bad_Konfig".Bad_Konfig[8].IO_Aus.LED_Einsetzen[2] THEN "FB_KP8_DB_5".KP8.LED[5] := 5; ELSE "FB_KP8_DB_5".KP8.LED[5] := 0; END_IF;
       IF "DB_Bad_Konfig".Bad_Konfig[8].IO_Aus.LED_Entnehmen[2] THEN
           IF "DB_Bad_Konfig".Bad_Konfig[8].IO_Aus.LED_Vorwarn[2] THEN "FB_KP8_DB_5".KP8.LED[1] := 4; ELSE "FB_KP8_DB_5".KP8.LED[1] := 5; END_IF;
       ELSE "FB_KP8_DB_5".KP8.LED[1] := 0; END_IF;
       IF "DB_Bad_Konfig".Bad_Konfig[8].IO_Aus.LED_Einsetzen[3] THEN "FB_KP8_DB_5".KP8.LED[4] := 5; ELSE "FB_KP8_DB_5".KP8.LED[4] := 0; END_IF;
       IF "DB_Bad_Konfig".Bad_Konfig[8].IO_Aus.LED_Entnehmen[3] THEN
           IF "DB_Bad_Konfig".Bad_Konfig[8].IO_Aus.LED_Vorwarn[3] THEN "FB_KP8_DB_5".KP8.LED[0] := 4; ELSE "FB_KP8_DB_5".KP8.LED[0] := 5; END_IF;
       ELSE "FB_KP8_DB_5".KP8.LED[0] := 0; END_IF;
       IF "DB_Bad_Konfig".Bad_Konfig[8].IO_Aus.LED_Heizung_Aktiv THEN "FB_KP8_DB_5".KP8.LED[3] := 4; ELSE "FB_KP8_DB_5".KP8.LED[3] := 0; END_IF;
       IF "DB_Bad_Konfig".Bad_Konfig[8].IO_Aus.LED_Stoerung THEN "FB_KP8_DB_5".KP8.LED[7] := 1; ELSE "FB_KP8_DB_5".KP8.LED[7] := 0; END_IF;
       IF "DB_Bad_Konfig".Bad_Konfig[12].IO_Aus.LED_Einsetzen[1] THEN "FB_KP8_DB_7".KP8.LED[6] := 5; ELSE "FB_KP8_DB_7".KP8.LED[6] := 0; END_IF;
       IF "DB_Bad_Konfig".Bad_Konfig[12].IO_Aus.LED_Entnehmen[1] THEN
           IF "DB_Bad_Konfig".Bad_Konfig[12].IO_Aus.LED_Vorwarn[1] THEN "FB_KP8_DB_7".KP8.LED[2] := 4; ELSE "FB_KP8_DB_7".KP8.LED[2] := 5; END_IF;
       ELSE "FB_KP8_DB_7".KP8.LED[2] := 0; END_IF;
       IF "DB_Bad_Konfig".Bad_Konfig[12].IO_Aus.LED_Einsetzen[2] THEN "FB_KP8_DB_7".KP8.LED[5] := 5; ELSE "FB_KP8_DB_7".KP8.LED[5] := 0; END_IF;
       IF "DB_Bad_Konfig".Bad_Konfig[12].IO_Aus.LED_Entnehmen[2] THEN
           IF "DB_Bad_Konfig".Bad_Konfig[12].IO_Aus.LED_Vorwarn[2] THEN "FB_KP8_DB_7".KP8.LED[1] := 4; ELSE "FB_KP8_DB_7".KP8.LED[1] := 5; END_IF;
       ELSE "FB_KP8_DB_7".KP8.LED[1] := 0; END_IF;
       IF "DB_Bad_Konfig".Bad_Konfig[12].IO_Aus.LED_Einsetzen[3] THEN "FB_KP8_DB_7".KP8.LED[4] := 5; ELSE "FB_KP8_DB_7".KP8.LED[4] := 0; END_IF;
       IF "DB_Bad_Konfig".Bad_Konfig[12].IO_Aus.LED_Entnehmen[3] THEN
           IF "DB_Bad_Konfig".Bad_Konfig[12].IO_Aus.LED_Vorwarn[3] THEN "FB_KP8_DB_7".KP8.LED[0] := 4; ELSE "FB_KP8_DB_7".KP8.LED[0] := 5; END_IF;
       ELSE "FB_KP8_DB_7".KP8.LED[0] := 0; END_IF;
       IF "DB_Bad_Konfig".Bad_Konfig[12].IO_Aus.LED_Heizung_Aktiv THEN "FB_KP8_DB_7".KP8.LED[3] := 4; ELSE "FB_KP8_DB_7".KP8.LED[3] := 0; END_IF;
       IF "DB_Bad_Konfig".Bad_Konfig[12].IO_Aus.LED_Stoerung THEN "FB_KP8_DB_7".KP8.LED[7] := 1; ELSE "FB_KP8_DB_7".KP8.LED[7] := 0; END_IF;
       IF "DB_Bad_Konfig".Bad_Konfig[13].IO_Aus.LED_Einsetzen[1] THEN "FB_KP8_DB_8".KP8.LED[6] := 5; ELSE "FB_KP8_DB_8".KP8.LED[6] := 0; END_IF;
       IF "DB_Bad_Konfig".Bad_Konfig[13].IO_Aus.LED_Entnehmen[1] THEN
           IF "DB_Bad_Konfig".Bad_Konfig[13].IO_Aus.LED_Vorwarn[1] THEN "FB_KP8_DB_8".KP8.LED[2] := 4; ELSE "FB_KP8_DB_8".KP8.LED[2] := 5; END_IF;
       ELSE "FB_KP8_DB_8".KP8.LED[2] := 0; END_IF;
       IF "DB_Bad_Konfig".Bad_Konfig[13].IO_Aus.LED_Einsetzen[2] THEN "FB_KP8_DB_8".KP8.LED[5] := 5; ELSE "FB_KP8_DB_8".KP8.LED[5] := 0; END_IF;
       IF "DB_Bad_Konfig".Bad_Konfig[13].IO_Aus.LED_Entnehmen[2] THEN
           IF "DB_Bad_Konfig".Bad_Konfig[13].IO_Aus.LED_Vorwarn[2] THEN "FB_KP8_DB_8".KP8.LED[1] := 4; ELSE "FB_KP8_DB_8".KP8.LED[1] := 5; END_IF;
       ELSE "FB_KP8_DB_8".KP8.LED[1] := 0; END_IF;
       IF "DB_Bad_Konfig".Bad_Konfig[13].IO_Aus.LED_Einsetzen[3] THEN "FB_KP8_DB_8".KP8.LED[4] := 5; ELSE "FB_KP8_DB_8".KP8.LED[4] := 0; END_IF;
       IF "DB_Bad_Konfig".Bad_Konfig[13].IO_Aus.LED_Entnehmen[3] THEN
           IF "DB_Bad_Konfig".Bad_Konfig[13].IO_Aus.LED_Vorwarn[3] THEN "FB_KP8_DB_8".KP8.LED[0] := 4; ELSE "FB_KP8_DB_8".KP8.LED[0] := 5; END_IF;
       ELSE "FB_KP8_DB_8".KP8.LED[0] := 0; END_IF;
       IF "DB_Bad_Konfig".Bad_Konfig[13].IO_Aus.LED_Heizung_Aktiv THEN "FB_KP8_DB_8".KP8.LED[3] := 4; ELSE "FB_KP8_DB_8".KP8.LED[3] := 0; END_IF;
       IF "DB_Bad_Konfig".Bad_Konfig[13].IO_Aus.LED_Stoerung THEN "FB_KP8_DB_8".KP8.LED[7] := 1; ELSE "FB_KP8_DB_8".KP8.LED[7] := 0; END_IF;
       IF "DB_Bad_Konfig".Bad_Konfig[14].IO_Aus.LED_Einsetzen[1] THEN "FB_KP8_DB_9".KP8.LED[6] := 5; ELSE "FB_KP8_DB_9".KP8.LED[6] := 0; END_IF;
       IF "DB_Bad_Konfig".Bad_Konfig[14].IO_Aus.LED_Entnehmen[1] THEN
           IF "DB_Bad_Konfig".Bad_Konfig[14].IO_Aus.LED_Vorwarn[1] THEN "FB_KP8_DB_9".KP8.LED[2] := 4; ELSE "FB_KP8_DB_9".KP8.LED[2] := 5; END_IF;
       ELSE "FB_KP8_DB_9".KP8.LED[2] := 0; END_IF;
       IF "DB_Bad_Konfig".Bad_Konfig[14].IO_Aus.LED_Einsetzen[2] THEN "FB_KP8_DB_9".KP8.LED[5] := 5; ELSE "FB_KP8_DB_9".KP8.LED[5] := 0; END_IF;
       IF "DB_Bad_Konfig".Bad_Konfig[14].IO_Aus.LED_Entnehmen[2] THEN
           IF "DB_Bad_Konfig".Bad_Konfig[14].IO_Aus.LED_Vorwarn[2] THEN "FB_KP8_DB_9".KP8.LED[1] := 4; ELSE "FB_KP8_DB_9".KP8.LED[1] := 5; END_IF;
       ELSE "FB_KP8_DB_9".KP8.LED[1] := 0; END_IF;
       IF "DB_Bad_Konfig".Bad_Konfig[14].IO_Aus.LED_Einsetzen[3] THEN "FB_KP8_DB_9".KP8.LED[4] := 5; ELSE "FB_KP8_DB_9".KP8.LED[4] := 0; END_IF;
       IF "DB_Bad_Konfig".Bad_Konfig[14].IO_Aus.LED_Entnehmen[3] THEN
           IF "DB_Bad_Konfig".Bad_Konfig[14].IO_Aus.LED_Vorwarn[3] THEN "FB_KP8_DB_9".KP8.LED[0] := 4; ELSE "FB_KP8_DB_9".KP8.LED[0] := 5; END_IF;
       ELSE "FB_KP8_DB_9".KP8.LED[0] := 0; END_IF;
       IF "DB_Bad_Konfig".Bad_Konfig[14].IO_Aus.LED_Heizung_Aktiv THEN "FB_KP8_DB_9".KP8.LED[3] := 4; ELSE "FB_KP8_DB_9".KP8.LED[3] := 0; END_IF;
       IF "DB_Bad_Konfig".Bad_Konfig[14].IO_Aus.LED_Stoerung THEN "FB_KP8_DB_9".KP8.LED[7] := 1; ELSE "FB_KP8_DB_9".KP8.LED[7] := 0; END_IF;
       IF "DB_Bad_Konfig".Bad_Konfig[18].IO_Aus.LED_Einsetzen[1] THEN "FB_KP8_DB_11".KP8.LED[6] := 5; ELSE "FB_KP8_DB_11".KP8.LED[6] := 0; END_IF;
       IF "DB_Bad_Konfig".Bad_Konfig[18].IO_Aus.LED_Entnehmen[1] THEN
           IF "DB_Bad_Konfig".Bad_Konfig[18].IO_Aus.LED_Vorwarn[1] THEN "FB_KP8_DB_11".KP8.LED[2] := 4; ELSE "FB_KP8_DB_11".KP8.LED[2] := 5; END_IF;
       ELSE "FB_KP8_DB_11".KP8.LED[2] := 0; END_IF;
       IF "DB_Bad_Konfig".Bad_Konfig[18].IO_Aus.LED_Einsetzen[2] THEN "FB_KP8_DB_11".KP8.LED[5] := 5; ELSE "FB_KP8_DB_11".KP8.LED[5] := 0; END_IF;
       IF "DB_Bad_Konfig".Bad_Konfig[18].IO_Aus.LED_Entnehmen[2] THEN
           IF "DB_Bad_Konfig".Bad_Konfig[18].IO_Aus.LED_Vorwarn[2] THEN "FB_KP8_DB_11".KP8.LED[1] := 4; ELSE "FB_KP8_DB_11".KP8.LED[1] := 5; END_IF;
       ELSE "FB_KP8_DB_11".KP8.LED[1] := 0; END_IF;
       IF "DB_Bad_Konfig".Bad_Konfig[18].IO_Aus.LED_Einsetzen[3] THEN "FB_KP8_DB_11".KP8.LED[4] := 5; ELSE "FB_KP8_DB_11".KP8.LED[4] := 0; END_IF;
       IF "DB_Bad_Konfig".Bad_Konfig[18].IO_Aus.LED_Entnehmen[3] THEN
           IF "DB_Bad_Konfig".Bad_Konfig[18].IO_Aus.LED_Vorwarn[3] THEN "FB_KP8_DB_11".KP8.LED[0] := 4; ELSE "FB_KP8_DB_11".KP8.LED[0] := 5; END_IF;
       ELSE "FB_KP8_DB_11".KP8.LED[0] := 0; END_IF;
       IF "DB_Bad_Konfig".Bad_Konfig[18].IO_Aus.LED_Heizung_Aktiv THEN "FB_KP8_DB_11".KP8.LED[3] := 4; ELSE "FB_KP8_DB_11".KP8.LED[3] := 0; END_IF;
       IF "DB_Bad_Konfig".Bad_Konfig[18].IO_Aus.LED_Stoerung THEN "FB_KP8_DB_11".KP8.LED[7] := 1; ELSE "FB_KP8_DB_11".KP8.LED[7] := 0; END_IF;
       IF "DB_Bad_Konfig".Bad_Konfig[19].IO_Aus.LED_Einsetzen[1] THEN "FB_KP8_DB_12".KP8.LED[6] := 5; ELSE "FB_KP8_DB_12".KP8.LED[6] := 0; END_IF;
       IF "DB_Bad_Konfig".Bad_Konfig[19].IO_Aus.LED_Entnehmen[1] THEN
           IF "DB_Bad_Konfig".Bad_Konfig[19].IO_Aus.LED_Vorwarn[1] THEN "FB_KP8_DB_12".KP8.LED[2] := 4; ELSE "FB_KP8_DB_12".KP8.LED[2] := 5; END_IF;
       ELSE "FB_KP8_DB_12".KP8.LED[2] := 0; END_IF;
       IF "DB_Bad_Konfig".Bad_Konfig[19].IO_Aus.LED_Einsetzen[2] THEN "FB_KP8_DB_12".KP8.LED[5] := 5; ELSE "FB_KP8_DB_12".KP8.LED[5] := 0; END_IF;
       IF "DB_Bad_Konfig".Bad_Konfig[19].IO_Aus.LED_Entnehmen[2] THEN
           IF "DB_Bad_Konfig".Bad_Konfig[19].IO_Aus.LED_Vorwarn[2] THEN "FB_KP8_DB_12".KP8.LED[1] := 4; ELSE "FB_KP8_DB_12".KP8.LED[1] := 5; END_IF;
       ELSE "FB_KP8_DB_12".KP8.LED[1] := 0; END_IF;
       IF "DB_Bad_Konfig".Bad_Konfig[19].IO_Aus.LED_Einsetzen[3] THEN "FB_KP8_DB_12".KP8.LED[4] := 5; ELSE "FB_KP8_DB_12".KP8.LED[4] := 0; END_IF;
       IF "DB_Bad_Konfig".Bad_Konfig[19].IO_Aus.LED_Entnehmen[3] THEN
           IF "DB_Bad_Konfig".Bad_Konfig[19].IO_Aus.LED_Vorwarn[3] THEN "FB_KP8_DB_12".KP8.LED[0] := 4; ELSE "FB_KP8_DB_12".KP8.LED[0] := 5; END_IF;
       ELSE "FB_KP8_DB_12".KP8.LED[0] := 0; END_IF;
       IF "DB_Bad_Konfig".Bad_Konfig[19].IO_Aus.LED_Heizung_Aktiv THEN "FB_KP8_DB_12".KP8.LED[3] := 4; ELSE "FB_KP8_DB_12".KP8.LED[3] := 0; END_IF;
       IF "DB_Bad_Konfig".Bad_Konfig[19].IO_Aus.LED_Stoerung THEN "FB_KP8_DB_12".KP8.LED[7] := 1; ELSE "FB_KP8_DB_12".KP8.LED[7] := 0; END_IF;
       IF "DB_Bad_Konfig".Bad_Konfig[21].IO_Aus.LED_Einsetzen[1] THEN "FB_KP8_DB_13".KP8.LED[6] := 5; ELSE "FB_KP8_DB_13".KP8.LED[6] := 0; END_IF;
       IF "DB_Bad_Konfig".Bad_Konfig[21].IO_Aus.LED_Entnehmen[1] THEN
           IF "DB_Bad_Konfig".Bad_Konfig[21].IO_Aus.LED_Vorwarn[1] THEN "FB_KP8_DB_13".KP8.LED[2] := 4; ELSE "FB_KP8_DB_13".KP8.LED[2] := 5; END_IF;
       ELSE "FB_KP8_DB_13".KP8.LED[2] := 0; END_IF;
       IF "DB_Bad_Konfig".Bad_Konfig[21].IO_Aus.LED_Einsetzen[2] THEN "FB_KP8_DB_13".KP8.LED[5] := 5; ELSE "FB_KP8_DB_13".KP8.LED[5] := 0; END_IF;
       IF "DB_Bad_Konfig".Bad_Konfig[21].IO_Aus.LED_Entnehmen[2] THEN
           IF "DB_Bad_Konfig".Bad_Konfig[21].IO_Aus.LED_Vorwarn[2] THEN "FB_KP8_DB_13".KP8.LED[1] := 4; ELSE "FB_KP8_DB_13".KP8.LED[1] := 5; END_IF;
       ELSE "FB_KP8_DB_13".KP8.LED[1] := 0; END_IF;
       IF "DB_Bad_Konfig".Bad_Konfig[21].IO_Aus.LED_Einsetzen[3] THEN "FB_KP8_DB_13".KP8.LED[4] := 5; ELSE "FB_KP8_DB_13".KP8.LED[4] := 0; END_IF;
       IF "DB_Bad_Konfig".Bad_Konfig[21].IO_Aus.LED_Entnehmen[3] THEN
           IF "DB_Bad_Konfig".Bad_Konfig[21].IO_Aus.LED_Vorwarn[3] THEN "FB_KP8_DB_13".KP8.LED[0] := 4; ELSE "FB_KP8_DB_13".KP8.LED[0] := 5; END_IF;
       ELSE "FB_KP8_DB_13".KP8.LED[0] := 0; END_IF;
       IF "DB_Bad_Konfig".Bad_Konfig[21].IO_Aus.LED_Heizung_Aktiv THEN "FB_KP8_DB_13".KP8.LED[3] := 4; ELSE "FB_KP8_DB_13".KP8.LED[3] := 0; END_IF;
       IF "DB_Bad_Konfig".Bad_Konfig[21].IO_Aus.LED_Stoerung THEN "FB_KP8_DB_13".KP8.LED[7] := 1; ELSE "FB_KP8_DB_13".KP8.LED[7] := 0; END_IF;
       IF "DB_Bad_Konfig".Bad_Konfig[26].IO_Aus.LED_Einsetzen[1] THEN "FB_KP8_DB_15".KP8.LED[6] := 5; ELSE "FB_KP8_DB_15".KP8.LED[6] := 0; END_IF;
       IF "DB_Bad_Konfig".Bad_Konfig[26].IO_Aus.LED_Entnehmen[1] THEN
           IF "DB_Bad_Konfig".Bad_Konfig[26].IO_Aus.LED_Vorwarn[1] THEN "FB_KP8_DB_15".KP8.LED[2] := 4; ELSE "FB_KP8_DB_15".KP8.LED[2] := 5; END_IF;
       ELSE "FB_KP8_DB_15".KP8.LED[2] := 0; END_IF;
       IF "DB_Bad_Konfig".Bad_Konfig[26].IO_Aus.LED_Einsetzen[2] THEN "FB_KP8_DB_15".KP8.LED[5] := 5; ELSE "FB_KP8_DB_15".KP8.LED[5] := 0; END_IF;
       IF "DB_Bad_Konfig".Bad_Konfig[26].IO_Aus.LED_Entnehmen[2] THEN
           IF "DB_Bad_Konfig".Bad_Konfig[26].IO_Aus.LED_Vorwarn[2] THEN "FB_KP8_DB_15".KP8.LED[1] := 4; ELSE "FB_KP8_DB_15".KP8.LED[1] := 5; END_IF;
       ELSE "FB_KP8_DB_15".KP8.LED[1] := 0; END_IF;
       IF "DB_Bad_Konfig".Bad_Konfig[26].IO_Aus.LED_Einsetzen[3] THEN "FB_KP8_DB_15".KP8.LED[4] := 5; ELSE "FB_KP8_DB_15".KP8.LED[4] := 0; END_IF;
       IF "DB_Bad_Konfig".Bad_Konfig[26].IO_Aus.LED_Entnehmen[3] THEN
           IF "DB_Bad_Konfig".Bad_Konfig[26].IO_Aus.LED_Vorwarn[3] THEN "FB_KP8_DB_15".KP8.LED[0] := 4; ELSE "FB_KP8_DB_15".KP8.LED[0] := 5; END_IF;
       ELSE "FB_KP8_DB_15".KP8.LED[0] := 0; END_IF;
       IF "DB_Bad_Konfig".Bad_Konfig[26].IO_Aus.LED_Heizung_Aktiv THEN "FB_KP8_DB_15".KP8.LED[3] := 4; ELSE "FB_KP8_DB_15".KP8.LED[3] := 0; END_IF;
       IF "DB_Bad_Konfig".Bad_Konfig[26].IO_Aus.LED_Stoerung THEN "FB_KP8_DB_15".KP8.LED[7] := 1; ELSE "FB_KP8_DB_15".KP8.LED[7] := 0; END_IF;
       IF "DB_Bad_Konfig".Bad_Konfig[30].IO_Aus.LED_Einsetzen[1] THEN "FB_KP8_DB_17".KP8.LED[6] := 5; ELSE "FB_KP8_DB_17".KP8.LED[6] := 0; END_IF;
       IF "DB_Bad_Konfig".Bad_Konfig[30].IO_Aus.LED_Entnehmen[1] THEN
           IF "DB_Bad_Konfig".Bad_Konfig[30].IO_Aus.LED_Vorwarn[1] THEN "FB_KP8_DB_17".KP8.LED[2] := 4; ELSE "FB_KP8_DB_17".KP8.LED[2] := 5; END_IF;
       ELSE "FB_KP8_DB_17".KP8.LED[2] := 0; END_IF;
       IF "DB_Bad_Konfig".Bad_Konfig[30].IO_Aus.LED_Einsetzen[2] THEN "FB_KP8_DB_17".KP8.LED[5] := 5; ELSE "FB_KP8_DB_17".KP8.LED[5] := 0; END_IF;
       IF "DB_Bad_Konfig".Bad_Konfig[30].IO_Aus.LED_Entnehmen[2] THEN
           IF "DB_Bad_Konfig".Bad_Konfig[30].IO_Aus.LED_Vorwarn[2] THEN "FB_KP8_DB_17".KP8.LED[1] := 4; ELSE "FB_KP8_DB_17".KP8.LED[1] := 5; END_IF;
       ELSE "FB_KP8_DB_17".KP8.LED[1] := 0; END_IF;
       IF "DB_Bad_Konfig".Bad_Konfig[30].IO_Aus.LED_Einsetzen[3] THEN "FB_KP8_DB_17".KP8.LED[4] := 5; ELSE "FB_KP8_DB_17".KP8.LED[4] := 0; END_IF;
       IF "DB_Bad_Konfig".Bad_Konfig[30].IO_Aus.LED_Entnehmen[3] THEN
           IF "DB_Bad_Konfig".Bad_Konfig[30].IO_Aus.LED_Vorwarn[3] THEN "FB_KP8_DB_17".KP8.LED[0] := 4; ELSE "FB_KP8_DB_17".KP8.LED[0] := 5; END_IF;
       ELSE "FB_KP8_DB_17".KP8.LED[0] := 0; END_IF;
       IF "DB_Bad_Konfig".Bad_Konfig[30].IO_Aus.LED_Heizung_Aktiv THEN "FB_KP8_DB_17".KP8.LED[3] := 4; ELSE "FB_KP8_DB_17".KP8.LED[3] := 0; END_IF;
       IF "DB_Bad_Konfig".Bad_Konfig[30].IO_Aus.LED_Stoerung THEN "FB_KP8_DB_17".KP8.LED[7] := 1; ELSE "FB_KP8_DB_17".KP8.LED[7] := 0; END_IF;
       IF "DB_Bad_Konfig".Bad_Konfig[31].IO_Aus.LED_Einsetzen[1] THEN "FB_KP8_DB_18".KP8.LED[6] := 5; ELSE "FB_KP8_DB_18".KP8.LED[6] := 0; END_IF;
       IF "DB_Bad_Konfig".Bad_Konfig[31].IO_Aus.LED_Entnehmen[1] THEN
           IF "DB_Bad_Konfig".Bad_Konfig[31].IO_Aus.LED_Vorwarn[1] THEN "FB_KP8_DB_18".KP8.LED[2] := 4; ELSE "FB_KP8_DB_18".KP8.LED[2] := 5; END_IF;
       ELSE "FB_KP8_DB_18".KP8.LED[2] := 0; END_IF;
       IF "DB_Bad_Konfig".Bad_Konfig[31].IO_Aus.LED_Einsetzen[2] THEN "FB_KP8_DB_18".KP8.LED[5] := 5; ELSE "FB_KP8_DB_18".KP8.LED[5] := 0; END_IF;
       IF "DB_Bad_Konfig".Bad_Konfig[31].IO_Aus.LED_Entnehmen[2] THEN
           IF "DB_Bad_Konfig".Bad_Konfig[31].IO_Aus.LED_Vorwarn[2] THEN "FB_KP8_DB_18".KP8.LED[1] := 4; ELSE "FB_KP8_DB_18".KP8.LED[1] := 5; END_IF;
       ELSE "FB_KP8_DB_18".KP8.LED[1] := 0; END_IF;
       IF "DB_Bad_Konfig".Bad_Konfig[31].IO_Aus.LED_Einsetzen[3] THEN "FB_KP8_DB_18".KP8.LED[4] := 5; ELSE "FB_KP8_DB_18".KP8.LED[4] := 0; END_IF;
       IF "DB_Bad_Konfig".Bad_Konfig[31].IO_Aus.LED_Entnehmen[3] THEN
           IF "DB_Bad_Konfig".Bad_Konfig[31].IO_Aus.LED_Vorwarn[3] THEN "FB_KP8_DB_18".KP8.LED[0] := 4; ELSE "FB_KP8_DB_18".KP8.LED[0] := 5; END_IF;
       ELSE "FB_KP8_DB_18".KP8.LED[0] := 0; END_IF;
       IF "DB_Bad_Konfig".Bad_Konfig[31].IO_Aus.LED_Heizung_Aktiv THEN "FB_KP8_DB_18".KP8.LED[3] := 4; ELSE "FB_KP8_DB_18".KP8.LED[3] := 0; END_IF;
       IF "DB_Bad_Konfig".Bad_Konfig[31].IO_Aus.LED_Stoerung THEN "FB_KP8_DB_18".KP8.LED[7] := 1; ELSE "FB_KP8_DB_18".KP8.LED[7] := 0; END_IF;
       IF "DB_Bad_Konfig".Bad_Konfig[35].IO_Aus.LED_Einsetzen[1] THEN "FB_KP8_DB_20".KP8.LED[6] := 5; ELSE "FB_KP8_DB_20".KP8.LED[6] := 0; END_IF;
       IF "DB_Bad_Konfig".Bad_Konfig[35].IO_Aus.LED_Entnehmen[1] THEN
           IF "DB_Bad_Konfig".Bad_Konfig[35].IO_Aus.LED_Vorwarn[1] THEN "FB_KP8_DB_20".KP8.LED[2] := 4; ELSE "FB_KP8_DB_20".KP8.LED[2] := 5; END_IF;
       ELSE "FB_KP8_DB_20".KP8.LED[2] := 0; END_IF;
       IF "DB_Bad_Konfig".Bad_Konfig[35].IO_Aus.LED_Einsetzen[2] THEN "FB_KP8_DB_20".KP8.LED[5] := 5; ELSE "FB_KP8_DB_20".KP8.LED[5] := 0; END_IF;
       IF "DB_Bad_Konfig".Bad_Konfig[35].IO_Aus.LED_Entnehmen[2] THEN
           IF "DB_Bad_Konfig".Bad_Konfig[35].IO_Aus.LED_Vorwarn[2] THEN "FB_KP8_DB_20".KP8.LED[1] := 4; ELSE "FB_KP8_DB_20".KP8.LED[1] := 5; END_IF;
       ELSE "FB_KP8_DB_20".KP8.LED[1] := 0; END_IF;
       IF "DB_Bad_Konfig".Bad_Konfig[35].IO_Aus.LED_Einsetzen[3] THEN "FB_KP8_DB_20".KP8.LED[4] := 5; ELSE "FB_KP8_DB_20".KP8.LED[4] := 0; END_IF;
       IF "DB_Bad_Konfig".Bad_Konfig[35].IO_Aus.LED_Entnehmen[3] THEN
           IF "DB_Bad_Konfig".Bad_Konfig[35].IO_Aus.LED_Vorwarn[3] THEN "FB_KP8_DB_20".KP8.LED[0] := 4; ELSE "FB_KP8_DB_20".KP8.LED[0] := 5; END_IF;
       ELSE "FB_KP8_DB_20".KP8.LED[0] := 0; END_IF;
       IF "DB_Bad_Konfig".Bad_Konfig[35].IO_Aus.LED_Heizung_Aktiv THEN "FB_KP8_DB_20".KP8.LED[3] := 4; ELSE "FB_KP8_DB_20".KP8.LED[3] := 0; END_IF;
       IF "DB_Bad_Konfig".Bad_Konfig[35].IO_Aus.LED_Stoerung THEN "FB_KP8_DB_20".KP8.LED[7] := 1; ELSE "FB_KP8_DB_20".KP8.LED[7] := 0; END_IF;
       IF "DB_Bad_Konfig".Bad_Konfig[36].IO_Aus.LED_Einsetzen[1] THEN "FB_KP8_DB_21".KP8.LED[6] := 5; ELSE "FB_KP8_DB_21".KP8.LED[6] := 0; END_IF;
       IF "DB_Bad_Konfig".Bad_Konfig[36].IO_Aus.LED_Entnehmen[1] THEN
           IF "DB_Bad_Konfig".Bad_Konfig[36].IO_Aus.LED_Vorwarn[1] THEN "FB_KP8_DB_21".KP8.LED[2] := 4; ELSE "FB_KP8_DB_21".KP8.LED[2] := 5; END_IF;
       ELSE "FB_KP8_DB_21".KP8.LED[2] := 0; END_IF;
       IF "DB_Bad_Konfig".Bad_Konfig[36].IO_Aus.LED_Einsetzen[2] THEN "FB_KP8_DB_21".KP8.LED[5] := 5; ELSE "FB_KP8_DB_21".KP8.LED[5] := 0; END_IF;
       IF "DB_Bad_Konfig".Bad_Konfig[36].IO_Aus.LED_Entnehmen[2] THEN
           IF "DB_Bad_Konfig".Bad_Konfig[36].IO_Aus.LED_Vorwarn[2] THEN "FB_KP8_DB_21".KP8.LED[1] := 4; ELSE "FB_KP8_DB_21".KP8.LED[1] := 5; END_IF;
       ELSE "FB_KP8_DB_21".KP8.LED[1] := 0; END_IF;
       IF "DB_Bad_Konfig".Bad_Konfig[36].IO_Aus.LED_Einsetzen[3] THEN "FB_KP8_DB_21".KP8.LED[4] := 5; ELSE "FB_KP8_DB_21".KP8.LED[4] := 0; END_IF;
       IF "DB_Bad_Konfig".Bad_Konfig[36].IO_Aus.LED_Entnehmen[3] THEN
           IF "DB_Bad_Konfig".Bad_Konfig[36].IO_Aus.LED_Vorwarn[3] THEN "FB_KP8_DB_21".KP8.LED[0] := 4; ELSE "FB_KP8_DB_21".KP8.LED[0] := 5; END_IF;
       ELSE "FB_KP8_DB_21".KP8.LED[0] := 0; END_IF;
       IF "DB_Bad_Konfig".Bad_Konfig[36].IO_Aus.LED_Heizung_Aktiv THEN "FB_KP8_DB_21".KP8.LED[3] := 4; ELSE "FB_KP8_DB_21".KP8.LED[3] := 0; END_IF;
       IF "DB_Bad_Konfig".Bad_Konfig[36].IO_Aus.LED_Stoerung THEN "FB_KP8_DB_21".KP8.LED[7] := 1; ELSE "FB_KP8_DB_21".KP8.LED[7] := 0; END_IF;
       IF "DB_Bad_Konfig".Bad_Konfig[40].IO_Aus.LED_Einsetzen[1] THEN "FB_KP8_DB_23".KP8.LED[6] := 5; ELSE "FB_KP8_DB_23".KP8.LED[6] := 0; END_IF;
       IF "DB_Bad_Konfig".Bad_Konfig[40].IO_Aus.LED_Entnehmen[1] THEN
           IF "DB_Bad_Konfig".Bad_Konfig[40].IO_Aus.LED_Vorwarn[1] THEN "FB_KP8_DB_23".KP8.LED[2] := 4; ELSE "FB_KP8_DB_23".KP8.LED[2] := 5; END_IF;
       ELSE "FB_KP8_DB_23".KP8.LED[2] := 0; END_IF;
       IF "DB_Bad_Konfig".Bad_Konfig[40].IO_Aus.LED_Einsetzen[2] THEN "FB_KP8_DB_23".KP8.LED[5] := 5; ELSE "FB_KP8_DB_23".KP8.LED[5] := 0; END_IF;
       IF "DB_Bad_Konfig".Bad_Konfig[40].IO_Aus.LED_Entnehmen[2] THEN
           IF "DB_Bad_Konfig".Bad_Konfig[40].IO_Aus.LED_Vorwarn[2] THEN "FB_KP8_DB_23".KP8.LED[1] := 4; ELSE "FB_KP8_DB_23".KP8.LED[1] := 5; END_IF;
       ELSE "FB_KP8_DB_23".KP8.LED[1] := 0; END_IF;
       IF "DB_Bad_Konfig".Bad_Konfig[40].IO_Aus.LED_Einsetzen[3] THEN "FB_KP8_DB_23".KP8.LED[4] := 5; ELSE "FB_KP8_DB_23".KP8.LED[4] := 0; END_IF;
       IF "DB_Bad_Konfig".Bad_Konfig[40].IO_Aus.LED_Entnehmen[3] THEN
           IF "DB_Bad_Konfig".Bad_Konfig[40].IO_Aus.LED_Vorwarn[3] THEN "FB_KP8_DB_23".KP8.LED[0] := 4; ELSE "FB_KP8_DB_23".KP8.LED[0] := 5; END_IF;
       ELSE "FB_KP8_DB_23".KP8.LED[0] := 0; END_IF;
       IF "DB_Bad_Konfig".Bad_Konfig[40].IO_Aus.LED_Heizung_Aktiv THEN "FB_KP8_DB_23".KP8.LED[3] := 4; ELSE "FB_KP8_DB_23".KP8.LED[3] := 0; END_IF;
       IF "DB_Bad_Konfig".Bad_Konfig[40].IO_Aus.LED_Stoerung THEN "FB_KP8_DB_23".KP8.LED[7] := 1; ELSE "FB_KP8_DB_23".KP8.LED[7] := 0; END_IF;
       IF "DB_Bad_Konfig".Bad_Konfig[41].IO_Aus.LED_Einsetzen[1] THEN "FB_KP8_DB_24".KP8.LED[6] := 5; ELSE "FB_KP8_DB_24".KP8.LED[6] := 0; END_IF;
       IF "DB_Bad_Konfig".Bad_Konfig[41].IO_Aus.LED_Entnehmen[1] THEN
           IF "DB_Bad_Konfig".Bad_Konfig[41].IO_Aus.LED_Vorwarn[1] THEN "FB_KP8_DB_24".KP8.LED[2] := 4; ELSE "FB_KP8_DB_24".KP8.LED[2] := 5; END_IF;
       ELSE "FB_KP8_DB_24".KP8.LED[2] := 0; END_IF;
       IF "DB_Bad_Konfig".Bad_Konfig[41].IO_Aus.LED_Einsetzen[2] THEN "FB_KP8_DB_24".KP8.LED[5] := 5; ELSE "FB_KP8_DB_24".KP8.LED[5] := 0; END_IF;
       IF "DB_Bad_Konfig".Bad_Konfig[41].IO_Aus.LED_Entnehmen[2] THEN
           IF "DB_Bad_Konfig".Bad_Konfig[41].IO_Aus.LED_Vorwarn[2] THEN "FB_KP8_DB_24".KP8.LED[1] := 4; ELSE "FB_KP8_DB_24".KP8.LED[1] := 5; END_IF;
       ELSE "FB_KP8_DB_24".KP8.LED[1] := 0; END_IF;
       IF "DB_Bad_Konfig".Bad_Konfig[41].IO_Aus.LED_Einsetzen[3] THEN "FB_KP8_DB_24".KP8.LED[4] := 5; ELSE "FB_KP8_DB_24".KP8.LED[4] := 0; END_IF;
       IF "DB_Bad_Konfig".Bad_Konfig[41].IO_Aus.LED_Entnehmen[3] THEN
           IF "DB_Bad_Konfig".Bad_Konfig[41].IO_Aus.LED_Vorwarn[3] THEN "FB_KP8_DB_24".KP8.LED[0] := 4; ELSE "FB_KP8_DB_24".KP8.LED[0] := 5; END_IF;
       ELSE "FB_KP8_DB_24".KP8.LED[0] := 0; END_IF;
       IF "DB_Bad_Konfig".Bad_Konfig[41].IO_Aus.LED_Heizung_Aktiv THEN "FB_KP8_DB_24".KP8.LED[3] := 4; ELSE "FB_KP8_DB_24".KP8.LED[3] := 0; END_IF;
       IF "DB_Bad_Konfig".Bad_Konfig[41].IO_Aus.LED_Stoerung THEN "FB_KP8_DB_24".KP8.LED[7] := 1; ELSE "FB_KP8_DB_24".KP8.LED[7] := 0; END_IF;
       IF "DB_Bad_Konfig".Bad_Konfig[45].IO_Aus.LED_Einsetzen[1] THEN "FB_KP8_DB_26".KP8.LED[6] := 5; ELSE "FB_KP8_DB_26".KP8.LED[6] := 0; END_IF;
       IF "DB_Bad_Konfig".Bad_Konfig[45].IO_Aus.LED_Entnehmen[1] THEN
           IF "DB_Bad_Konfig".Bad_Konfig[45].IO_Aus.LED_Vorwarn[1] THEN "FB_KP8_DB_26".KP8.LED[2] := 4; ELSE "FB_KP8_DB_26".KP8.LED[2] := 5; END_IF;
       ELSE "FB_KP8_DB_26".KP8.LED[2] := 0; END_IF;
       IF "DB_Bad_Konfig".Bad_Konfig[45].IO_Aus.LED_Einsetzen[2] THEN "FB_KP8_DB_26".KP8.LED[5] := 5; ELSE "FB_KP8_DB_26".KP8.LED[5] := 0; END_IF;
       IF "DB_Bad_Konfig".Bad_Konfig[45].IO_Aus.LED_Entnehmen[2] THEN
           IF "DB_Bad_Konfig".Bad_Konfig[45].IO_Aus.LED_Vorwarn[2] THEN "FB_KP8_DB_26".KP8.LED[1] := 4; ELSE "FB_KP8_DB_26".KP8.LED[1] := 5; END_IF;
       ELSE "FB_KP8_DB_26".KP8.LED[1] := 0; END_IF;
       IF "DB_Bad_Konfig".Bad_Konfig[45].IO_Aus.LED_Einsetzen[3] THEN "FB_KP8_DB_26".KP8.LED[4] := 5; ELSE "FB_KP8_DB_26".KP8.LED[4] := 0; END_IF;
       IF "DB_Bad_Konfig".Bad_Konfig[45].IO_Aus.LED_Entnehmen[3] THEN
           IF "DB_Bad_Konfig".Bad_Konfig[45].IO_Aus.LED_Vorwarn[3] THEN "FB_KP8_DB_26".KP8.LED[0] := 4; ELSE "FB_KP8_DB_26".KP8.LED[0] := 5; END_IF;
       ELSE "FB_KP8_DB_26".KP8.LED[0] := 0; END_IF;
       IF "DB_Bad_Konfig".Bad_Konfig[45].IO_Aus.LED_Heizung_Aktiv THEN "FB_KP8_DB_26".KP8.LED[3] := 4; ELSE "FB_KP8_DB_26".KP8.LED[3] := 0; END_IF;
       IF "DB_Bad_Konfig".Bad_Konfig[45].IO_Aus.LED_Stoerung THEN "FB_KP8_DB_26".KP8.LED[7] := 1; ELSE "FB_KP8_DB_26".KP8.LED[7] := 0; END_IF;
       IF "DB_Bad_Konfig".Bad_Konfig[46].IO_Aus.LED_Einsetzen[1] THEN "FB_KP8_DB_27".KP8.LED[6] := 5; ELSE "FB_KP8_DB_27".KP8.LED[6] := 0; END_IF;
       IF "DB_Bad_Konfig".Bad_Konfig[46].IO_Aus.LED_Entnehmen[1] THEN
           IF "DB_Bad_Konfig".Bad_Konfig[46].IO_Aus.LED_Vorwarn[1] THEN "FB_KP8_DB_27".KP8.LED[2] := 4; ELSE "FB_KP8_DB_27".KP8.LED[2] := 5; END_IF;
       ELSE "FB_KP8_DB_27".KP8.LED[2] := 0; END_IF;
       IF "DB_Bad_Konfig".Bad_Konfig[46].IO_Aus.LED_Einsetzen[2] THEN "FB_KP8_DB_27".KP8.LED[5] := 5; ELSE "FB_KP8_DB_27".KP8.LED[5] := 0; END_IF;
       IF "DB_Bad_Konfig".Bad_Konfig[46].IO_Aus.LED_Entnehmen[2] THEN
           IF "DB_Bad_Konfig".Bad_Konfig[46].IO_Aus.LED_Vorwarn[2] THEN "FB_KP8_DB_27".KP8.LED[1] := 4; ELSE "FB_KP8_DB_27".KP8.LED[1] := 5; END_IF;
       ELSE "FB_KP8_DB_27".KP8.LED[1] := 0; END_IF;
       IF "DB_Bad_Konfig".Bad_Konfig[46].IO_Aus.LED_Einsetzen[3] THEN "FB_KP8_DB_27".KP8.LED[4] := 5; ELSE "FB_KP8_DB_27".KP8.LED[4] := 0; END_IF;
       IF "DB_Bad_Konfig".Bad_Konfig[46].IO_Aus.LED_Entnehmen[3] THEN
           IF "DB_Bad_Konfig".Bad_Konfig[46].IO_Aus.LED_Vorwarn[3] THEN "FB_KP8_DB_27".KP8.LED[0] := 4; ELSE "FB_KP8_DB_27".KP8.LED[0] := 5; END_IF;
       ELSE "FB_KP8_DB_27".KP8.LED[0] := 0; END_IF;
       IF "DB_Bad_Konfig".Bad_Konfig[46].IO_Aus.LED_Heizung_Aktiv THEN "FB_KP8_DB_27".KP8.LED[3] := 4; ELSE "FB_KP8_DB_27".KP8.LED[3] := 0; END_IF;
       IF "DB_Bad_Konfig".Bad_Konfig[46].IO_Aus.LED_Stoerung THEN "FB_KP8_DB_27".KP8.LED[7] := 1; ELSE "FB_KP8_DB_27".KP8.LED[7] := 0; END_IF;
       IF "DB_Bad_Konfig".Bad_Konfig[25].IO_Aus.LED_Einsetzen[1] THEN "FB_KP8_DB_28".KP8.LED[6] := 5; ELSE "FB_KP8_DB_28".KP8.LED[6] := 0; END_IF;
       IF "DB_Bad_Konfig".Bad_Konfig[25].IO_Aus.LED_Entnehmen[1] THEN
           IF "DB_Bad_Konfig".Bad_Konfig[25].IO_Aus.LED_Vorwarn[1] THEN "FB_KP8_DB_28".KP8.LED[2] := 4; ELSE "FB_KP8_DB_28".KP8.LED[2] := 5; END_IF;
       ELSE "FB_KP8_DB_28".KP8.LED[2] := 0; END_IF;
       IF "DB_Bad_Konfig".Bad_Konfig[25].IO_Aus.LED_Einsetzen[2] THEN "FB_KP8_DB_28".KP8.LED[5] := 5; ELSE "FB_KP8_DB_28".KP8.LED[5] := 0; END_IF;
       IF "DB_Bad_Konfig".Bad_Konfig[25].IO_Aus.LED_Entnehmen[2] THEN
           IF "DB_Bad_Konfig".Bad_Konfig[25].IO_Aus.LED_Vorwarn[2] THEN "FB_KP8_DB_28".KP8.LED[1] := 4; ELSE "FB_KP8_DB_28".KP8.LED[1] := 5; END_IF;
       ELSE "FB_KP8_DB_28".KP8.LED[1] := 0; END_IF;
       IF "DB_Bad_Konfig".Bad_Konfig[25].IO_Aus.LED_Einsetzen[3] THEN "FB_KP8_DB_28".KP8.LED[4] := 5; ELSE "FB_KP8_DB_28".KP8.LED[4] := 0; END_IF;
       IF "DB_Bad_Konfig".Bad_Konfig[25].IO_Aus.LED_Entnehmen[3] THEN
           IF "DB_Bad_Konfig".Bad_Konfig[25].IO_Aus.LED_Vorwarn[3] THEN "FB_KP8_DB_28".KP8.LED[0] := 4; ELSE "FB_KP8_DB_28".KP8.LED[0] := 5; END_IF;
       ELSE "FB_KP8_DB_28".KP8.LED[0] := 0; END_IF;
       IF "DB_Bad_Konfig".Bad_Konfig[25].IO_Aus.LED_Heizung_Aktiv THEN "FB_KP8_DB_28".KP8.LED[3] := 4; ELSE "FB_KP8_DB_28".KP8.LED[3] := 0; END_IF;
       IF "DB_Bad_Konfig".Bad_Konfig[25].IO_Aus.LED_Stoerung THEN "FB_KP8_DB_28".KP8.LED[7] := 1; ELSE "FB_KP8_DB_28".KP8.LED[7] := 0; END_IF;
       #pw := "DB_Bad_Konfig".Bad_Konfig[4].IO_Aus.Prio_Einsetzen_WT;
       "FB_KP8_DB_3".KP8.LED[4] := 0;
       IF (#pw >= 1) AND (#pw <= 3) THEN
           IF "DB_Bad_Konfig".Bad_Konfig[4].IO_Aus.LED_Einsetzen[#pw] THEN "FB_KP8_DB_3".KP8.LED[4] := 5; END_IF;
       END_IF;
       #pw := "DB_Bad_Konfig".Bad_Konfig[4].IO_Aus.Prio_Entnehmen_WT;
       "FB_KP8_DB_3".KP8.LED[0] := 0;
       IF (#pw >= 1) AND (#pw <= 3) THEN
           IF "DB_Bad_Konfig".Bad_Konfig[4].IO_Aus.LED_Entnehmen[#pw] THEN
               IF "DB_Bad_Konfig".Bad_Konfig[4].IO_Aus.LED_Vorwarn[#pw] THEN "FB_KP8_DB_3".KP8.LED[0] := 4; ELSE "FB_KP8_DB_3".KP8.LED[0] := 5; END_IF;
           END_IF;
       END_IF;
       #pw := "DB_Bad_Konfig".Bad_Konfig[5].IO_Aus.Prio_Einsetzen_WT;
       "FB_KP8_DB_3".KP8.LED[5] := 0;
       IF (#pw >= 1) AND (#pw <= 3) THEN
           IF "DB_Bad_Konfig".Bad_Konfig[5].IO_Aus.LED_Einsetzen[#pw] THEN "FB_KP8_DB_3".KP8.LED[5] := 5; END_IF;
       END_IF;
       #pw := "DB_Bad_Konfig".Bad_Konfig[5].IO_Aus.Prio_Entnehmen_WT;
       "FB_KP8_DB_3".KP8.LED[1] := 0;
       IF (#pw >= 1) AND (#pw <= 3) THEN
           IF "DB_Bad_Konfig".Bad_Konfig[5].IO_Aus.LED_Entnehmen[#pw] THEN
               IF "DB_Bad_Konfig".Bad_Konfig[5].IO_Aus.LED_Vorwarn[#pw] THEN "FB_KP8_DB_3".KP8.LED[1] := 4; ELSE "FB_KP8_DB_3".KP8.LED[1] := 5; END_IF;
           END_IF;
       END_IF;
       #pw := "DB_Bad_Konfig".Bad_Konfig[6].IO_Aus.Prio_Einsetzen_WT;
       "FB_KP8_DB_3".KP8.LED[6] := 0;
       IF (#pw >= 1) AND (#pw <= 3) THEN
           IF "DB_Bad_Konfig".Bad_Konfig[6].IO_Aus.LED_Einsetzen[#pw] THEN "FB_KP8_DB_3".KP8.LED[6] := 5; END_IF;
       END_IF;
       #pw := "DB_Bad_Konfig".Bad_Konfig[6].IO_Aus.Prio_Entnehmen_WT;
       "FB_KP8_DB_3".KP8.LED[2] := 0;
       IF (#pw >= 1) AND (#pw <= 3) THEN
           IF "DB_Bad_Konfig".Bad_Konfig[6].IO_Aus.LED_Entnehmen[#pw] THEN
               IF "DB_Bad_Konfig".Bad_Konfig[6].IO_Aus.LED_Vorwarn[#pw] THEN "FB_KP8_DB_3".KP8.LED[2] := 4; ELSE "FB_KP8_DB_3".KP8.LED[2] := 5; END_IF;
           END_IF;
       END_IF;
       IF "DB_Bad_Konfig".Bad_Konfig[4].IO_Aus.LED_Heizung_Aktiv OR "DB_Bad_Konfig".Bad_Konfig[5].IO_Aus.LED_Heizung_Aktiv OR "DB_Bad_Konfig".Bad_Konfig[6].IO_Aus.LED_Heizung_Aktiv THEN "FB_KP8_DB_3".KP8.LED[3] := 4; ELSE "FB_KP8_DB_3".KP8.LED[3] := 0; END_IF;
       IF "DB_Bad_Konfig".Bad_Konfig[4].IO_Aus.LED_Stoerung OR "DB_Bad_Konfig".Bad_Konfig[5].IO_Aus.LED_Stoerung OR "DB_Bad_Konfig".Bad_Konfig[6].IO_Aus.LED_Stoerung THEN "FB_KP8_DB_3".KP8.LED[7] := 1; ELSE "FB_KP8_DB_3".KP8.LED[7] := 0; END_IF;
       #pw := "DB_Bad_Konfig".Bad_Konfig[9].IO_Aus.Prio_Einsetzen_WT;
       "FB_KP8_DB_6".KP8.LED[4] := 0;
       IF (#pw >= 1) AND (#pw <= 3) THEN
           IF "DB_Bad_Konfig".Bad_Konfig[9].IO_Aus.LED_Einsetzen[#pw] THEN "FB_KP8_DB_6".KP8.LED[4] := 5; END_IF;
       END_IF;
       #pw := "DB_Bad_Konfig".Bad_Konfig[9].IO_Aus.Prio_Entnehmen_WT;
       "FB_KP8_DB_6".KP8.LED[0] := 0;
       IF (#pw >= 1) AND (#pw <= 3) THEN
           IF "DB_Bad_Konfig".Bad_Konfig[9].IO_Aus.LED_Entnehmen[#pw] THEN
               IF "DB_Bad_Konfig".Bad_Konfig[9].IO_Aus.LED_Vorwarn[#pw] THEN "FB_KP8_DB_6".KP8.LED[0] := 4; ELSE "FB_KP8_DB_6".KP8.LED[0] := 5; END_IF;
           END_IF;
       END_IF;
       #pw := "DB_Bad_Konfig".Bad_Konfig[10].IO_Aus.Prio_Einsetzen_WT;
       "FB_KP8_DB_6".KP8.LED[5] := 0;
       IF (#pw >= 1) AND (#pw <= 3) THEN
           IF "DB_Bad_Konfig".Bad_Konfig[10].IO_Aus.LED_Einsetzen[#pw] THEN "FB_KP8_DB_6".KP8.LED[5] := 5; END_IF;
       END_IF;
       #pw := "DB_Bad_Konfig".Bad_Konfig[10].IO_Aus.Prio_Entnehmen_WT;
       "FB_KP8_DB_6".KP8.LED[1] := 0;
       IF (#pw >= 1) AND (#pw <= 3) THEN
           IF "DB_Bad_Konfig".Bad_Konfig[10].IO_Aus.LED_Entnehmen[#pw] THEN
               IF "DB_Bad_Konfig".Bad_Konfig[10].IO_Aus.LED_Vorwarn[#pw] THEN "FB_KP8_DB_6".KP8.LED[1] := 4; ELSE "FB_KP8_DB_6".KP8.LED[1] := 5; END_IF;
           END_IF;
       END_IF;
       #pw := "DB_Bad_Konfig".Bad_Konfig[11].IO_Aus.Prio_Einsetzen_WT;
       "FB_KP8_DB_6".KP8.LED[6] := 0;
       IF (#pw >= 1) AND (#pw <= 3) THEN
           IF "DB_Bad_Konfig".Bad_Konfig[11].IO_Aus.LED_Einsetzen[#pw] THEN "FB_KP8_DB_6".KP8.LED[6] := 5; END_IF;
       END_IF;
       #pw := "DB_Bad_Konfig".Bad_Konfig[11].IO_Aus.Prio_Entnehmen_WT;
       "FB_KP8_DB_6".KP8.LED[2] := 0;
       IF (#pw >= 1) AND (#pw <= 3) THEN
           IF "DB_Bad_Konfig".Bad_Konfig[11].IO_Aus.LED_Entnehmen[#pw] THEN
               IF "DB_Bad_Konfig".Bad_Konfig[11].IO_Aus.LED_Vorwarn[#pw] THEN "FB_KP8_DB_6".KP8.LED[2] := 4; ELSE "FB_KP8_DB_6".KP8.LED[2] := 5; END_IF;
           END_IF;
       END_IF;
       IF "DB_Bad_Konfig".Bad_Konfig[9].IO_Aus.LED_Heizung_Aktiv OR "DB_Bad_Konfig".Bad_Konfig[10].IO_Aus.LED_Heizung_Aktiv OR "DB_Bad_Konfig".Bad_Konfig[11].IO_Aus.LED_Heizung_Aktiv THEN "FB_KP8_DB_6".KP8.LED[3] := 4; ELSE "FB_KP8_DB_6".KP8.LED[3] := 0; END_IF;
       IF "DB_Bad_Konfig".Bad_Konfig[9].IO_Aus.LED_Stoerung OR "DB_Bad_Konfig".Bad_Konfig[10].IO_Aus.LED_Stoerung OR "DB_Bad_Konfig".Bad_Konfig[11].IO_Aus.LED_Stoerung THEN "FB_KP8_DB_6".KP8.LED[7] := 1; ELSE "FB_KP8_DB_6".KP8.LED[7] := 0; END_IF;
       #pw := "DB_Bad_Konfig".Bad_Konfig[15].IO_Aus.Prio_Einsetzen_WT;
       "FB_KP8_DB_10".KP8.LED[4] := 0;
       IF (#pw >= 1) AND (#pw <= 3) THEN
           IF "DB_Bad_Konfig".Bad_Konfig[15].IO_Aus.LED_Einsetzen[#pw] THEN "FB_KP8_DB_10".KP8.LED[4] := 5; END_IF;
       END_IF;
       #pw := "DB_Bad_Konfig".Bad_Konfig[15].IO_Aus.Prio_Entnehmen_WT;
       "FB_KP8_DB_10".KP8.LED[0] := 0;
       IF (#pw >= 1) AND (#pw <= 3) THEN
           IF "DB_Bad_Konfig".Bad_Konfig[15].IO_Aus.LED_Entnehmen[#pw] THEN
               IF "DB_Bad_Konfig".Bad_Konfig[15].IO_Aus.LED_Vorwarn[#pw] THEN "FB_KP8_DB_10".KP8.LED[0] := 4; ELSE "FB_KP8_DB_10".KP8.LED[0] := 5; END_IF;
           END_IF;
       END_IF;
       #pw := "DB_Bad_Konfig".Bad_Konfig[16].IO_Aus.Prio_Einsetzen_WT;
       "FB_KP8_DB_10".KP8.LED[5] := 0;
       IF (#pw >= 1) AND (#pw <= 3) THEN
           IF "DB_Bad_Konfig".Bad_Konfig[16].IO_Aus.LED_Einsetzen[#pw] THEN "FB_KP8_DB_10".KP8.LED[5] := 5; END_IF;
       END_IF;
       #pw := "DB_Bad_Konfig".Bad_Konfig[16].IO_Aus.Prio_Entnehmen_WT;
       "FB_KP8_DB_10".KP8.LED[1] := 0;
       IF (#pw >= 1) AND (#pw <= 3) THEN
           IF "DB_Bad_Konfig".Bad_Konfig[16].IO_Aus.LED_Entnehmen[#pw] THEN
               IF "DB_Bad_Konfig".Bad_Konfig[16].IO_Aus.LED_Vorwarn[#pw] THEN "FB_KP8_DB_10".KP8.LED[1] := 4; ELSE "FB_KP8_DB_10".KP8.LED[1] := 5; END_IF;
           END_IF;
       END_IF;
       #pw := "DB_Bad_Konfig".Bad_Konfig[17].IO_Aus.Prio_Einsetzen_WT;
       "FB_KP8_DB_10".KP8.LED[6] := 0;
       IF (#pw >= 1) AND (#pw <= 3) THEN
           IF "DB_Bad_Konfig".Bad_Konfig[17].IO_Aus.LED_Einsetzen[#pw] THEN "FB_KP8_DB_10".KP8.LED[6] := 5; END_IF;
       END_IF;
       #pw := "DB_Bad_Konfig".Bad_Konfig[17].IO_Aus.Prio_Entnehmen_WT;
       "FB_KP8_DB_10".KP8.LED[2] := 0;
       IF (#pw >= 1) AND (#pw <= 3) THEN
           IF "DB_Bad_Konfig".Bad_Konfig[17].IO_Aus.LED_Entnehmen[#pw] THEN
               IF "DB_Bad_Konfig".Bad_Konfig[17].IO_Aus.LED_Vorwarn[#pw] THEN "FB_KP8_DB_10".KP8.LED[2] := 4; ELSE "FB_KP8_DB_10".KP8.LED[2] := 5; END_IF;
           END_IF;
       END_IF;
       IF "DB_Bad_Konfig".Bad_Konfig[15].IO_Aus.LED_Heizung_Aktiv OR "DB_Bad_Konfig".Bad_Konfig[16].IO_Aus.LED_Heizung_Aktiv OR "DB_Bad_Konfig".Bad_Konfig[17].IO_Aus.LED_Heizung_Aktiv THEN "FB_KP8_DB_10".KP8.LED[3] := 4; ELSE "FB_KP8_DB_10".KP8.LED[3] := 0; END_IF;
       IF "DB_Bad_Konfig".Bad_Konfig[15].IO_Aus.LED_Stoerung OR "DB_Bad_Konfig".Bad_Konfig[16].IO_Aus.LED_Stoerung OR "DB_Bad_Konfig".Bad_Konfig[17].IO_Aus.LED_Stoerung THEN "FB_KP8_DB_10".KP8.LED[7] := 1; ELSE "FB_KP8_DB_10".KP8.LED[7] := 0; END_IF;
       #pw := "DB_Bad_Konfig".Bad_Konfig[22].IO_Aus.Prio_Einsetzen_WT;
       "FB_KP8_DB_14".KP8.LED[4] := 0;
       IF (#pw >= 1) AND (#pw <= 3) THEN
           IF "DB_Bad_Konfig".Bad_Konfig[22].IO_Aus.LED_Einsetzen[#pw] THEN "FB_KP8_DB_14".KP8.LED[4] := 5; END_IF;
       END_IF;
       #pw := "DB_Bad_Konfig".Bad_Konfig[22].IO_Aus.Prio_Entnehmen_WT;
       "FB_KP8_DB_14".KP8.LED[0] := 0;
       IF (#pw >= 1) AND (#pw <= 3) THEN
           IF "DB_Bad_Konfig".Bad_Konfig[22].IO_Aus.LED_Entnehmen[#pw] THEN
               IF "DB_Bad_Konfig".Bad_Konfig[22].IO_Aus.LED_Vorwarn[#pw] THEN "FB_KP8_DB_14".KP8.LED[0] := 4; ELSE "FB_KP8_DB_14".KP8.LED[0] := 5; END_IF;
           END_IF;
       END_IF;
       #pw := "DB_Bad_Konfig".Bad_Konfig[23].IO_Aus.Prio_Einsetzen_WT;
       "FB_KP8_DB_14".KP8.LED[5] := 0;
       IF (#pw >= 1) AND (#pw <= 3) THEN
           IF "DB_Bad_Konfig".Bad_Konfig[23].IO_Aus.LED_Einsetzen[#pw] THEN "FB_KP8_DB_14".KP8.LED[5] := 5; END_IF;
       END_IF;
       #pw := "DB_Bad_Konfig".Bad_Konfig[23].IO_Aus.Prio_Entnehmen_WT;
       "FB_KP8_DB_14".KP8.LED[1] := 0;
       IF (#pw >= 1) AND (#pw <= 3) THEN
           IF "DB_Bad_Konfig".Bad_Konfig[23].IO_Aus.LED_Entnehmen[#pw] THEN
               IF "DB_Bad_Konfig".Bad_Konfig[23].IO_Aus.LED_Vorwarn[#pw] THEN "FB_KP8_DB_14".KP8.LED[1] := 4; ELSE "FB_KP8_DB_14".KP8.LED[1] := 5; END_IF;
           END_IF;
       END_IF;
       #pw := "DB_Bad_Konfig".Bad_Konfig[24].IO_Aus.Prio_Einsetzen_WT;
       "FB_KP8_DB_14".KP8.LED[6] := 0;
       IF (#pw >= 1) AND (#pw <= 3) THEN
           IF "DB_Bad_Konfig".Bad_Konfig[24].IO_Aus.LED_Einsetzen[#pw] THEN "FB_KP8_DB_14".KP8.LED[6] := 5; END_IF;
       END_IF;
       #pw := "DB_Bad_Konfig".Bad_Konfig[24].IO_Aus.Prio_Entnehmen_WT;
       "FB_KP8_DB_14".KP8.LED[2] := 0;
       IF (#pw >= 1) AND (#pw <= 3) THEN
           IF "DB_Bad_Konfig".Bad_Konfig[24].IO_Aus.LED_Entnehmen[#pw] THEN
               IF "DB_Bad_Konfig".Bad_Konfig[24].IO_Aus.LED_Vorwarn[#pw] THEN "FB_KP8_DB_14".KP8.LED[2] := 4; ELSE "FB_KP8_DB_14".KP8.LED[2] := 5; END_IF;
           END_IF;
       END_IF;
       IF "DB_Bad_Konfig".Bad_Konfig[22].IO_Aus.LED_Heizung_Aktiv OR "DB_Bad_Konfig".Bad_Konfig[23].IO_Aus.LED_Heizung_Aktiv OR "DB_Bad_Konfig".Bad_Konfig[24].IO_Aus.LED_Heizung_Aktiv THEN "FB_KP8_DB_14".KP8.LED[3] := 4; ELSE "FB_KP8_DB_14".KP8.LED[3] := 0; END_IF;
       IF "DB_Bad_Konfig".Bad_Konfig[22].IO_Aus.LED_Stoerung OR "DB_Bad_Konfig".Bad_Konfig[23].IO_Aus.LED_Stoerung OR "DB_Bad_Konfig".Bad_Konfig[24].IO_Aus.LED_Stoerung THEN "FB_KP8_DB_14".KP8.LED[7] := 1; ELSE "FB_KP8_DB_14".KP8.LED[7] := 0; END_IF;
       #pw := "DB_Bad_Konfig".Bad_Konfig[27].IO_Aus.Prio_Einsetzen_WT;
       "FB_KP8_DB_16".KP8.LED[4] := 0;
       IF (#pw >= 1) AND (#pw <= 3) THEN
           IF "DB_Bad_Konfig".Bad_Konfig[27].IO_Aus.LED_Einsetzen[#pw] THEN "FB_KP8_DB_16".KP8.LED[4] := 5; END_IF;
       END_IF;
       #pw := "DB_Bad_Konfig".Bad_Konfig[27].IO_Aus.Prio_Entnehmen_WT;
       "FB_KP8_DB_16".KP8.LED[0] := 0;
       IF (#pw >= 1) AND (#pw <= 3) THEN
           IF "DB_Bad_Konfig".Bad_Konfig[27].IO_Aus.LED_Entnehmen[#pw] THEN
               IF "DB_Bad_Konfig".Bad_Konfig[27].IO_Aus.LED_Vorwarn[#pw] THEN "FB_KP8_DB_16".KP8.LED[0] := 4; ELSE "FB_KP8_DB_16".KP8.LED[0] := 5; END_IF;
           END_IF;
       END_IF;
       #pw := "DB_Bad_Konfig".Bad_Konfig[28].IO_Aus.Prio_Einsetzen_WT;
       "FB_KP8_DB_16".KP8.LED[5] := 0;
       IF (#pw >= 1) AND (#pw <= 3) THEN
           IF "DB_Bad_Konfig".Bad_Konfig[28].IO_Aus.LED_Einsetzen[#pw] THEN "FB_KP8_DB_16".KP8.LED[5] := 5; END_IF;
       END_IF;
       #pw := "DB_Bad_Konfig".Bad_Konfig[28].IO_Aus.Prio_Entnehmen_WT;
       "FB_KP8_DB_16".KP8.LED[1] := 0;
       IF (#pw >= 1) AND (#pw <= 3) THEN
           IF "DB_Bad_Konfig".Bad_Konfig[28].IO_Aus.LED_Entnehmen[#pw] THEN
               IF "DB_Bad_Konfig".Bad_Konfig[28].IO_Aus.LED_Vorwarn[#pw] THEN "FB_KP8_DB_16".KP8.LED[1] := 4; ELSE "FB_KP8_DB_16".KP8.LED[1] := 5; END_IF;
           END_IF;
       END_IF;
       #pw := "DB_Bad_Konfig".Bad_Konfig[29].IO_Aus.Prio_Einsetzen_WT;
       "FB_KP8_DB_16".KP8.LED[6] := 0;
       IF (#pw >= 1) AND (#pw <= 3) THEN
           IF "DB_Bad_Konfig".Bad_Konfig[29].IO_Aus.LED_Einsetzen[#pw] THEN "FB_KP8_DB_16".KP8.LED[6] := 5; END_IF;
       END_IF;
       #pw := "DB_Bad_Konfig".Bad_Konfig[29].IO_Aus.Prio_Entnehmen_WT;
       "FB_KP8_DB_16".KP8.LED[2] := 0;
       IF (#pw >= 1) AND (#pw <= 3) THEN
           IF "DB_Bad_Konfig".Bad_Konfig[29].IO_Aus.LED_Entnehmen[#pw] THEN
               IF "DB_Bad_Konfig".Bad_Konfig[29].IO_Aus.LED_Vorwarn[#pw] THEN "FB_KP8_DB_16".KP8.LED[2] := 4; ELSE "FB_KP8_DB_16".KP8.LED[2] := 5; END_IF;
           END_IF;
       END_IF;
       IF "DB_Bad_Konfig".Bad_Konfig[27].IO_Aus.LED_Heizung_Aktiv OR "DB_Bad_Konfig".Bad_Konfig[28].IO_Aus.LED_Heizung_Aktiv OR "DB_Bad_Konfig".Bad_Konfig[29].IO_Aus.LED_Heizung_Aktiv THEN "FB_KP8_DB_16".KP8.LED[3] := 4; ELSE "FB_KP8_DB_16".KP8.LED[3] := 0; END_IF;
       IF "DB_Bad_Konfig".Bad_Konfig[27].IO_Aus.LED_Stoerung OR "DB_Bad_Konfig".Bad_Konfig[28].IO_Aus.LED_Stoerung OR "DB_Bad_Konfig".Bad_Konfig[29].IO_Aus.LED_Stoerung THEN "FB_KP8_DB_16".KP8.LED[7] := 1; ELSE "FB_KP8_DB_16".KP8.LED[7] := 0; END_IF;
       #pw := "DB_Bad_Konfig".Bad_Konfig[32].IO_Aus.Prio_Einsetzen_WT;
       "FB_KP8_DB_19".KP8.LED[4] := 0;
       IF (#pw >= 1) AND (#pw <= 3) THEN
           IF "DB_Bad_Konfig".Bad_Konfig[32].IO_Aus.LED_Einsetzen[#pw] THEN "FB_KP8_DB_19".KP8.LED[4] := 5; END_IF;
       END_IF;
       #pw := "DB_Bad_Konfig".Bad_Konfig[32].IO_Aus.Prio_Entnehmen_WT;
       "FB_KP8_DB_19".KP8.LED[0] := 0;
       IF (#pw >= 1) AND (#pw <= 3) THEN
           IF "DB_Bad_Konfig".Bad_Konfig[32].IO_Aus.LED_Entnehmen[#pw] THEN
               IF "DB_Bad_Konfig".Bad_Konfig[32].IO_Aus.LED_Vorwarn[#pw] THEN "FB_KP8_DB_19".KP8.LED[0] := 4; ELSE "FB_KP8_DB_19".KP8.LED[0] := 5; END_IF;
           END_IF;
       END_IF;
       #pw := "DB_Bad_Konfig".Bad_Konfig[33].IO_Aus.Prio_Einsetzen_WT;
       "FB_KP8_DB_19".KP8.LED[5] := 0;
       IF (#pw >= 1) AND (#pw <= 3) THEN
           IF "DB_Bad_Konfig".Bad_Konfig[33].IO_Aus.LED_Einsetzen[#pw] THEN "FB_KP8_DB_19".KP8.LED[5] := 5; END_IF;
       END_IF;
       #pw := "DB_Bad_Konfig".Bad_Konfig[33].IO_Aus.Prio_Entnehmen_WT;
       "FB_KP8_DB_19".KP8.LED[1] := 0;
       IF (#pw >= 1) AND (#pw <= 3) THEN
           IF "DB_Bad_Konfig".Bad_Konfig[33].IO_Aus.LED_Entnehmen[#pw] THEN
               IF "DB_Bad_Konfig".Bad_Konfig[33].IO_Aus.LED_Vorwarn[#pw] THEN "FB_KP8_DB_19".KP8.LED[1] := 4; ELSE "FB_KP8_DB_19".KP8.LED[1] := 5; END_IF;
           END_IF;
       END_IF;
       #pw := "DB_Bad_Konfig".Bad_Konfig[34].IO_Aus.Prio_Einsetzen_WT;
       "FB_KP8_DB_19".KP8.LED[6] := 0;
       IF (#pw >= 1) AND (#pw <= 3) THEN
           IF "DB_Bad_Konfig".Bad_Konfig[34].IO_Aus.LED_Einsetzen[#pw] THEN "FB_KP8_DB_19".KP8.LED[6] := 5; END_IF;
       END_IF;
       #pw := "DB_Bad_Konfig".Bad_Konfig[34].IO_Aus.Prio_Entnehmen_WT;
       "FB_KP8_DB_19".KP8.LED[2] := 0;
       IF (#pw >= 1) AND (#pw <= 3) THEN
           IF "DB_Bad_Konfig".Bad_Konfig[34].IO_Aus.LED_Entnehmen[#pw] THEN
               IF "DB_Bad_Konfig".Bad_Konfig[34].IO_Aus.LED_Vorwarn[#pw] THEN "FB_KP8_DB_19".KP8.LED[2] := 4; ELSE "FB_KP8_DB_19".KP8.LED[2] := 5; END_IF;
           END_IF;
       END_IF;
       IF "DB_Bad_Konfig".Bad_Konfig[32].IO_Aus.LED_Heizung_Aktiv OR "DB_Bad_Konfig".Bad_Konfig[33].IO_Aus.LED_Heizung_Aktiv OR "DB_Bad_Konfig".Bad_Konfig[34].IO_Aus.LED_Heizung_Aktiv THEN "FB_KP8_DB_19".KP8.LED[3] := 4; ELSE "FB_KP8_DB_19".KP8.LED[3] := 0; END_IF;
       IF "DB_Bad_Konfig".Bad_Konfig[32].IO_Aus.LED_Stoerung OR "DB_Bad_Konfig".Bad_Konfig[33].IO_Aus.LED_Stoerung OR "DB_Bad_Konfig".Bad_Konfig[34].IO_Aus.LED_Stoerung THEN "FB_KP8_DB_19".KP8.LED[7] := 1; ELSE "FB_KP8_DB_19".KP8.LED[7] := 0; END_IF;
       #pw := "DB_Bad_Konfig".Bad_Konfig[37].IO_Aus.Prio_Einsetzen_WT;
       "FB_KP8_DB_22".KP8.LED[4] := 0;
       IF (#pw >= 1) AND (#pw <= 3) THEN
           IF "DB_Bad_Konfig".Bad_Konfig[37].IO_Aus.LED_Einsetzen[#pw] THEN "FB_KP8_DB_22".KP8.LED[4] := 5; END_IF;
       END_IF;
       #pw := "DB_Bad_Konfig".Bad_Konfig[37].IO_Aus.Prio_Entnehmen_WT;
       "FB_KP8_DB_22".KP8.LED[0] := 0;
       IF (#pw >= 1) AND (#pw <= 3) THEN
           IF "DB_Bad_Konfig".Bad_Konfig[37].IO_Aus.LED_Entnehmen[#pw] THEN
               IF "DB_Bad_Konfig".Bad_Konfig[37].IO_Aus.LED_Vorwarn[#pw] THEN "FB_KP8_DB_22".KP8.LED[0] := 4; ELSE "FB_KP8_DB_22".KP8.LED[0] := 5; END_IF;
           END_IF;
       END_IF;
       #pw := "DB_Bad_Konfig".Bad_Konfig[38].IO_Aus.Prio_Einsetzen_WT;
       "FB_KP8_DB_22".KP8.LED[5] := 0;
       IF (#pw >= 1) AND (#pw <= 3) THEN
           IF "DB_Bad_Konfig".Bad_Konfig[38].IO_Aus.LED_Einsetzen[#pw] THEN "FB_KP8_DB_22".KP8.LED[5] := 5; END_IF;
       END_IF;
       #pw := "DB_Bad_Konfig".Bad_Konfig[38].IO_Aus.Prio_Entnehmen_WT;
       "FB_KP8_DB_22".KP8.LED[1] := 0;
       IF (#pw >= 1) AND (#pw <= 3) THEN
           IF "DB_Bad_Konfig".Bad_Konfig[38].IO_Aus.LED_Entnehmen[#pw] THEN
               IF "DB_Bad_Konfig".Bad_Konfig[38].IO_Aus.LED_Vorwarn[#pw] THEN "FB_KP8_DB_22".KP8.LED[1] := 4; ELSE "FB_KP8_DB_22".KP8.LED[1] := 5; END_IF;
           END_IF;
       END_IF;
       #pw := "DB_Bad_Konfig".Bad_Konfig[39].IO_Aus.Prio_Einsetzen_WT;
       "FB_KP8_DB_22".KP8.LED[6] := 0;
       IF (#pw >= 1) AND (#pw <= 3) THEN
           IF "DB_Bad_Konfig".Bad_Konfig[39].IO_Aus.LED_Einsetzen[#pw] THEN "FB_KP8_DB_22".KP8.LED[6] := 5; END_IF;
       END_IF;
       #pw := "DB_Bad_Konfig".Bad_Konfig[39].IO_Aus.Prio_Entnehmen_WT;
       "FB_KP8_DB_22".KP8.LED[2] := 0;
       IF (#pw >= 1) AND (#pw <= 3) THEN
           IF "DB_Bad_Konfig".Bad_Konfig[39].IO_Aus.LED_Entnehmen[#pw] THEN
               IF "DB_Bad_Konfig".Bad_Konfig[39].IO_Aus.LED_Vorwarn[#pw] THEN "FB_KP8_DB_22".KP8.LED[2] := 4; ELSE "FB_KP8_DB_22".KP8.LED[2] := 5; END_IF;
           END_IF;
       END_IF;
       IF "DB_Bad_Konfig".Bad_Konfig[37].IO_Aus.LED_Heizung_Aktiv OR "DB_Bad_Konfig".Bad_Konfig[38].IO_Aus.LED_Heizung_Aktiv OR "DB_Bad_Konfig".Bad_Konfig[39].IO_Aus.LED_Heizung_Aktiv THEN "FB_KP8_DB_22".KP8.LED[3] := 4; ELSE "FB_KP8_DB_22".KP8.LED[3] := 0; END_IF;
       IF "DB_Bad_Konfig".Bad_Konfig[37].IO_Aus.LED_Stoerung OR "DB_Bad_Konfig".Bad_Konfig[38].IO_Aus.LED_Stoerung OR "DB_Bad_Konfig".Bad_Konfig[39].IO_Aus.LED_Stoerung THEN "FB_KP8_DB_22".KP8.LED[7] := 1; ELSE "FB_KP8_DB_22".KP8.LED[7] := 0; END_IF;
       #pw := "DB_Bad_Konfig".Bad_Konfig[42].IO_Aus.Prio_Einsetzen_WT;
       "FB_KP8_DB_25".KP8.LED[4] := 0;
       IF (#pw >= 1) AND (#pw <= 3) THEN
           IF "DB_Bad_Konfig".Bad_Konfig[42].IO_Aus.LED_Einsetzen[#pw] THEN "FB_KP8_DB_25".KP8.LED[4] := 5; END_IF;
       END_IF;
       #pw := "DB_Bad_Konfig".Bad_Konfig[42].IO_Aus.Prio_Entnehmen_WT;
       "FB_KP8_DB_25".KP8.LED[0] := 0;
       IF (#pw >= 1) AND (#pw <= 3) THEN
           IF "DB_Bad_Konfig".Bad_Konfig[42].IO_Aus.LED_Entnehmen[#pw] THEN
               IF "DB_Bad_Konfig".Bad_Konfig[42].IO_Aus.LED_Vorwarn[#pw] THEN "FB_KP8_DB_25".KP8.LED[0] := 4; ELSE "FB_KP8_DB_25".KP8.LED[0] := 5; END_IF;
           END_IF;
       END_IF;
       #pw := "DB_Bad_Konfig".Bad_Konfig[43].IO_Aus.Prio_Einsetzen_WT;
       "FB_KP8_DB_25".KP8.LED[5] := 0;
       IF (#pw >= 1) AND (#pw <= 3) THEN
           IF "DB_Bad_Konfig".Bad_Konfig[43].IO_Aus.LED_Einsetzen[#pw] THEN "FB_KP8_DB_25".KP8.LED[5] := 5; END_IF;
       END_IF;
       #pw := "DB_Bad_Konfig".Bad_Konfig[43].IO_Aus.Prio_Entnehmen_WT;
       "FB_KP8_DB_25".KP8.LED[1] := 0;
       IF (#pw >= 1) AND (#pw <= 3) THEN
           IF "DB_Bad_Konfig".Bad_Konfig[43].IO_Aus.LED_Entnehmen[#pw] THEN
               IF "DB_Bad_Konfig".Bad_Konfig[43].IO_Aus.LED_Vorwarn[#pw] THEN "FB_KP8_DB_25".KP8.LED[1] := 4; ELSE "FB_KP8_DB_25".KP8.LED[1] := 5; END_IF;
           END_IF;
       END_IF;
       #pw := "DB_Bad_Konfig".Bad_Konfig[44].IO_Aus.Prio_Einsetzen_WT;
       "FB_KP8_DB_25".KP8.LED[6] := 0;
       IF (#pw >= 1) AND (#pw <= 3) THEN
           IF "DB_Bad_Konfig".Bad_Konfig[44].IO_Aus.LED_Einsetzen[#pw] THEN "FB_KP8_DB_25".KP8.LED[6] := 5; END_IF;
       END_IF;
       #pw := "DB_Bad_Konfig".Bad_Konfig[44].IO_Aus.Prio_Entnehmen_WT;
       "FB_KP8_DB_25".KP8.LED[2] := 0;
       IF (#pw >= 1) AND (#pw <= 3) THEN
           IF "DB_Bad_Konfig".Bad_Konfig[44].IO_Aus.LED_Entnehmen[#pw] THEN
               IF "DB_Bad_Konfig".Bad_Konfig[44].IO_Aus.LED_Vorwarn[#pw] THEN "FB_KP8_DB_25".KP8.LED[2] := 4; ELSE "FB_KP8_DB_25".KP8.LED[2] := 5; END_IF;
           END_IF;
       END_IF;
       IF "DB_Bad_Konfig".Bad_Konfig[42].IO_Aus.LED_Heizung_Aktiv OR "DB_Bad_Konfig".Bad_Konfig[43].IO_Aus.LED_Heizung_Aktiv OR "DB_Bad_Konfig".Bad_Konfig[44].IO_Aus.LED_Heizung_Aktiv THEN "FB_KP8_DB_25".KP8.LED[3] := 4; ELSE "FB_KP8_DB_25".KP8.LED[3] := 0; END_IF;
       IF "DB_Bad_Konfig".Bad_Konfig[42].IO_Aus.LED_Stoerung OR "DB_Bad_Konfig".Bad_Konfig[43].IO_Aus.LED_Stoerung OR "DB_Bad_Konfig".Bad_Konfig[44].IO_Aus.LED_Stoerung THEN "FB_KP8_DB_25".KP8.LED[7] := 1; ELSE "FB_KP8_DB_25".KP8.LED[7] := 0; END_IF;

       // Peripherie-Ausgaenge
       "Pumpe Bad 8"      := "DB_Bad_Konfig".Bad_Konfig[8].IO_Aus.Pumpe;
       "Pumpe Bad 12"     := "DB_Bad_Konfig".Bad_Konfig[12].IO_Aus.Pumpe;
       "Pumpe Bad 14"     := "DB_Bad_Konfig".Bad_Konfig[14].IO_Aus.Pumpe;
       "Pumpe Bad 18"     := "DB_Bad_Konfig".Bad_Konfig[18].IO_Aus.Pumpe;
       "Pumpe Bad 19"     := "DB_Bad_Konfig".Bad_Konfig[19].IO_Aus.Pumpe;
       "Pumpe Bad 21"     := "DB_Bad_Konfig".Bad_Konfig[21].IO_Aus.Pumpe;
       // Bad 25: Netzschuetz + FU
       "Netzschuetz Pumpe Bad 25"   := "DB_Bad_Konfig".Bad_Konfig[25].IO_Aus.Pumpe_FU_Netzschuetz;
       "FU Pumpe Freigabe"          := "DB_Bad_Konfig".Bad_Konfig[25].IO_Aus.Pumpe_FU_Freigabe;
       "Reset FU Pumpe"             := "DB_Bad_Konfig".Bad_Konfig[25].IO_Aus.Pumpe_FU_Reset;
       "Pumpen_FU_Steuerwert"       := INT_TO_WORD(REAL_TO_INT("DB_Bad_Konfig".Bad_Konfig[25].Pumpe_FU_Soll * 276.48));
       "Pumpe Bad 26"     := "DB_Bad_Konfig".Bad_Konfig[26].IO_Aus.Pumpe;
       "Pumpe Bad 31"     := "DB_Bad_Konfig".Bad_Konfig[31].IO_Aus.Pumpe;
       "Pumpe Bad 41"     := "DB_Bad_Konfig".Bad_Konfig[41].IO_Aus.Pumpe;
       "Pumpe Bad 45"     := "DB_Bad_Konfig".Bad_Konfig[45].IO_Aus.Pumpe;

       // Heizungen
       "Regelung Heizung Bad 7"           := "DB_Bad_Konfig".Bad_Konfig[7].IO_Aus.Heizung_1_Regelung;
       "Sicherheitsschuetz Heizung Bad 7"  := "DB_Bad_Konfig".Bad_Konfig[7].IO_Aus.Heizung_1_Sicherheit;
       "Regelung Heizung Bad 8"           := "DB_Bad_Konfig".Bad_Konfig[8].IO_Aus.Heizung_1_Regelung;
       "Sicherheitsschuetz Heizung Bad 8"  := "DB_Bad_Konfig".Bad_Konfig[8].IO_Aus.Heizung_1_Sicherheit;
       "Regelung Heizung Bad 12"          := "DB_Bad_Konfig".Bad_Konfig[12].IO_Aus.Heizung_1_Regelung;
       "Sicherheitsschuetz Heizung Bad 12" := "DB_Bad_Konfig".Bad_Konfig[12].IO_Aus.Heizung_1_Sicherheit;
       "Regelung Heizung 1 Bad 25"        := "DB_Bad_Konfig".Bad_Konfig[25].IO_Aus.Heizung_1_Regelung;
       "Regelung Heizung 2 Bad 25"        := "DB_Bad_Konfig".Bad_Konfig[25].IO_Aus.Heizung_2_Regelung;
       "Sicherheitsschuetze Heizung 1 + 2 Bad 25" := "DB_Bad_Konfig".Bad_Konfig[25].IO_Aus.Heizung_1_Sicherheit OR "DB_Bad_Konfig".Bad_Konfig[25].IO_Aus.Heizung_2_Sicherheit;
       "Regelung Heizung Bad 36"          := "DB_Bad_Konfig".Bad_Konfig[36].IO_Aus.Heizung_1_Regelung;
       "Sicherheitsschuetz Heizung Bad 36" := "DB_Bad_Konfig".Bad_Konfig[36].IO_Aus.Heizung_1_Sicherheit;
       "Regelung Heizung Bad 40"          := "DB_Bad_Konfig".Bad_Konfig[40].IO_Aus.Heizung_1_Regelung;
       "Sicherheitsschuetz Heizung Bad 40" := "DB_Bad_Konfig".Bad_Konfig[40].IO_Aus.Heizung_1_Sicherheit;
       "Regelung Heizung Bad 46"          := "DB_Bad_Konfig".Bad_Konfig[46].IO_Aus.Heizung_1_Regelung;
       "Sicherheitsschuetz Heizung Bad 46" := "DB_Bad_Konfig".Bad_Konfig[46].IO_Aus.Heizung_1_Sicherheit;
       "Freigabe Ultraschall Pos. 8"  := "DB_Bad_Konfig".Bad_Konfig[8].IO_Aus.Ultraschall_Freigabe;
       "Freigabe Ultraschall Pos. 12" := "DB_Bad_Konfig".Bad_Konfig[12].IO_Aus.Ultraschall_Freigabe;

       // Warenbewegung Bad 25 (X=WB2, Y=WB1 physisch)
       "Warenbewegung 1 Bad 25 Netzschuetz"  := "DB_Bad_Konfig".Bad_Konfig[25].Warenbewegung_Y_Soll > 0.0;
       "Warenbewegung 1 Bad 25 Freigabe FU" := "DB_Bad_Konfig".Bad_Konfig[25].Warenbewegung_Y_Soll > 0.0;
       "Warenbewegung 1 Bad 25 Reset FU"    := "DB_Bad_Konfig".Bad_Konfig[25].WB1_Reset;
       "Warenbewegung 2 Bad 25 Netzschuetz"  := "DB_Bad_Konfig".Bad_Konfig[25].Warenbewegung_X_Soll > 0.0;
       "Warenbewegung 2 Bad 25 Freigabe FU" := "DB_Bad_Konfig".Bad_Konfig[25].Warenbewegung_X_Soll > 0.0;
       "Warenbewegung 2 Bad 25 Reset FU"    := "DB_Bad_Konfig".Bad_Konfig[25].WB2_Reset;
       "Warenbewegung 1 Bad 25 Sollwert FU" := INT_TO_WORD(REAL_TO_INT("DB_Bad_Konfig".Bad_Konfig[25].Warenbewegung_Y_Soll * 276.48));
       "Warenbewegung 2 Bad 25 Sollwert FU" := INT_TO_WORD(REAL_TO_INT("DB_Bad_Konfig".Bad_Konfig[25].Warenbewegung_X_Soll * 276.48));

       // Hupe
       #hupe_sammel := FALSE;
       FOR #b := 1 TO "c_Anzahl_Bad" DO IF "DB_Bad_Konfig".Bad_Konfig[#b].Hupe THEN #hupe_sammel := TRUE; END_IF; END_FOR;
       "Masch.Leuchte 1 Anlage Hupe" := #hupe_sammel;
   END_IF;
END_FUNCTION

FUNCTION "FC_KP8_Override" : Void   // FC4, SCL
{ S7_Optimized_Access := 'TRUE' }
VERSION : 0.1
// stored: AutoNumber true, IsIECCheckEnabled false, SetENOAutomatically false, UDAEnableTagReadback false
   VAR_INPUT
      Lampentest : Bool;
      Blink_Takt : Bool;
   END_VAR
   VAR_TEMP
      i : Int;
      led_val : USInt;
   END_VAR
BEGIN

